{region 'Documentation'}
(*!
<summary>Number of observations from the latest subject call.</summary>
*)
{endregion}
{attribute 'monitoring' := 'call'}
PROPERTY PUBLIC HookCount : UINT //! Number of observations from the latest subject call.
GET // PUBLIC
HookCount := FHookCount;
END_GET
END_PROPERTY

{region 'Documentation'}
(*!
<summary>Combines base startability with the scenario release.</summary>
*)
{endregion}
{attribute 'monitoring' := 'call'}
PROPERTY PUBLIC IsReady : BOOL //! Combines base startability with the scenario release.
GET // PUBLIC
IsReady := SUPER^.IsReady AND Ready;
END_GET
END_PROPERTY

{region 'Documentation'}
(*!
<summary>
Records activation, supports a controlled cleanup failure and waits for the explicit completion release.
</summary>
*)
{endregion}
METHOD PROTECTED ProcessAbort
VAR_INPUT
    Enable : BOOL; //! Phase permission supplied by the owning Test Case; FALSE does not authorize progression, while observation may continue.
END_VAR
RecordHook(Hook := E_LifecycleHook.Abort,
    Enabled := Enable);
IF NOT Enable THEN
    RETURN;
END_IF;
IF AbortError THEN
    Error(Message := 'Controlled abort failure.');
END_IF;
IF AbortCompleted THEN
    CompleteAbort();
END_IF;
END_METHOD

{region 'Documentation'}
(*!
<summary>Calls both real Assertions even when disabled to consume their reset requests.</summary>
*)
{endregion}
METHOD PROTECTED ProcessAssertions
VAR_INPUT
    Enable : BOOL; //! Phase permission supplied by the owning Test Case; FALSE does not authorize progression, while observation may continue.
END_VAR
RecordHook(Hook := E_LifecycleHook.Assertions,
    Enabled := Enable);
FAssertion(Enable := Enable,
    State := State,
    IN := AssertionCondition);
FReferenceAssertion(Enable := Enable,
    State := State,
    IN := TRUE);
END_METHOD

{region 'Documentation'}
(*!
<summary>Supplies controlled target observations and explicit multi-stage completion.</summary>
*)
{endregion}
METHOD PROTECTED ProcessPreparations
VAR_INPUT
    Enable : BOOL; //! Phase permission supplied by the owning Test Case; FALSE does not authorize progression, while observation may continue.
END_VAR
RecordHook(Hook := E_LifecycleHook.Preparations,
    Enabled := Enable);
// Emulate the concrete application's combined observation without another Preparation FB.
// The Sequencer has already run; explicit completion below can still transition immediately.
UpdatePreparationStatus(Ready := TRUE,
    Running := Enable AND NOT PreparationTargetReached,
    Completed := PreparationTargetReached,
    HasError := PreparationError);
IF NOT Enable THEN
    RETURN;
END_IF;

IF AdvancePreparation THEN
    NextPreparationState();
ELSIF FinishPreparations THEN
    CompletePreparations();
END_IF;
END_METHOD

{region 'Documentation'}
(*!
<summary>Resets both real Assertions and completes only on the explicit fixture release.</summary>
*)
{endregion}
METHOD PROTECTED ProcessReset
RecordHook(Hook := E_LifecycleHook.Reset,
    Enabled := TRUE);
FAssertion.Reset();
FReferenceAssertion.Reset();
// Deliberately allow Error followed by CompleteReset in the same call.
// The base must preserve Error and choose finalization instead of a successful Idle result.
IF ResetError THEN
    Error(Message := 'Controlled reset failure.');
END_IF;
IF ResetCompleted THEN
    CompleteReset();
END_IF;
END_METHOD

{region 'Documentation'}
(*!
<summary>Advances or completes only when enabled and explicitly instructed.</summary>
*)
{endregion}
METHOD PROTECTED ProcessTests
VAR_INPUT
    Enable : BOOL; //! Phase permission supplied by the owning Test Case; FALSE does not authorize progression, while observation may continue.
END_VAR
RecordHook(Hook := E_LifecycleHook.Tests,
    Enabled := Enable);
IF NOT Enable THEN
    RETURN;
END_IF;

// Use the real base API for error and transition stimulus; never assign the subject state directly.
IF TestError THEN
    Error(Message := 'Controlled test failure.');
    RETURN;
END_IF;
IF AdvanceTest THEN
    NextTestState();
ELSIF FinishTests THEN
    CompleteTests();
END_IF;
END_METHOD

{region 'Documentation'}
(*!
<summary>Appends one hook-entry observation with bounded storage and explicit overflow reporting.</summary>
*)
{endregion}
METHOD PRIVATE RecordHook
VAR_INPUT
    Hook : E_LifecycleHook; //! Hook being entered; appended to the bounded per-call trace.
    Enabled : BOOL; //! Hook permission recorded together with the current entry state.
END_VAR
IF FHookCount >= HookCapacity THEN
    FTraceOverflow := TRUE;
    RETURN;
END_IF;

FHookCount := FHookCount + 1;
FHooks[FHookCount].Hook := Hook;
FHooks[FHookCount].State := State;
FHooks[FHookCount].Enabled := Enabled;
END_METHOD

{region 'Documentation'}
(*!
<summary>Reports a call exceeding the bounded hook trace.</summary>
*)
{endregion}
{attribute 'monitoring' := 'call'}
PROPERTY PUBLIC TraceOverflow : BOOL //! Reports a call exceeding the bounded hook trace.
GET // PUBLIC
TraceOverflow := FTraceOverflow;
END_GET
END_PROPERTY

END_FUNCTION_BLOCK

// ---- SelfTests/TestCases/TestSuite_TestCaseLifecycle/Test_LifecycleWithoutPreparation.TcPOU
{region 'Documentation'}
(*!
<summary>Checks initial passivity, parent Reset, resource readiness and explicit single-state completion.</summary>
*)
{endregion}
FUNCTION_BLOCK Test_LifecycleWithoutPreparation EXTENDS TestCaseLifecycleTestBase

SUPER^();

{region 'Documentation'}
(*!
<summary>Defines independent per-call stimuli and expected lifecycle/hook observations.</summary>
*)
{endregion}
METHOD PROTECTED ConfigureScenario
FSubjectPreparationCount := 0;
FSubjectTestCount := 1;
FStepCount := 11;

{region "01 - Initialized but awaiting Reset"}
// After successful Initialize, remain Uninitialized until the parent requests Reset.
FSteps[1].ExpectedState := E_State.Uninitialized;
FSteps[1].ExpectedResult := E_Result.NotEvaluated;
FSteps[1].ExpectedReady := FALSE;
FSteps[1].ExpectedPassedCount := 0;
FSteps[1].ExpectedFailedCount := 0;
FSteps[1].ExpectedHookCount := 5;
FSteps[1].ExpectedHooks[1].Hook := E_LifecycleHook.Abort;
FSteps[1].ExpectedHooks[1].State := E_State.Uninitialized;
FSteps[1].ExpectedHooks[1].Enabled := FALSE;
FSteps[1].ExpectedHooks[2].Hook := E_LifecycleHook.Preparations;
FSteps[1].ExpectedHooks[2].State := E_State.Uninitialized;
FSteps[1].ExpectedHooks[2].Enabled := FALSE;
FSteps[1].ExpectedHooks[3].Hook := E_LifecycleHook.Tests;
FSteps[1].ExpectedHooks[3].State := E_State.Uninitialized;
FSteps[1].ExpectedHooks[3].Enabled := FALSE;
FSteps[1].ExpectedHooks[4].Hook := E_LifecycleHook.Assertions;
FSteps[1].ExpectedHooks[4].State := E_State.Uninitialized;
FSteps[1].ExpectedHooks[4].Enabled := FALSE;
FSteps[1].ExpectedHooks[5].Hook := E_LifecycleHook.Aggregate;
FSteps[1].ExpectedHooks[5].State := E_State.Uninitialized;
FSteps[1].ExpectedHooks[5].Enabled := TRUE;
{endregion}

{region "02 - Start cannot bypass Reset"}
// Start alone must not bypass the initial Reset requirement.
FSteps[2].RequestStart := TRUE;
FSteps[2].ExpectedState := E_State.Uninitialized;
FSteps[2].ExpectedResult := E_Result.NotEvaluated;
FSteps[2].ExpectedReady := FALSE;
FSteps[2].ExpectedPassedCount := 0;
FSteps[2].ExpectedFailedCount := 0;
FSteps[2].ExpectedHookCount := 5;
FSteps[2].ExpectedHooks[1].Hook := E_LifecycleHook.Abort;
FSteps[2].ExpectedHooks[1].State := E_State.Uninitialized;
FSteps[2].ExpectedHooks[1].Enabled := FALSE;
FSteps[2].ExpectedHooks[2].Hook := E_LifecycleHook.Preparations;
FSteps[2].ExpectedHooks[2].State := E_State.Uninitialized;
FSteps[2].ExpectedHooks[2].Enabled := FALSE;
FSteps[2].ExpectedHooks[3].Hook := E_LifecycleHook.Tests;
FSteps[2].ExpectedHooks[3].State := E_State.Uninitialized;
FSteps[2].ExpectedHooks[3].Enabled := FALSE;
FSteps[2].ExpectedHooks[4].Hook := E_LifecycleHook.Assertions;
FSteps[2].ExpectedHooks[4].State := E_State.Uninitialized;
FSteps[2].ExpectedHooks[4].Enabled := FALSE;
FSteps[2].ExpectedHooks[5].Hook := E_LifecycleHook.Aggregate;
FSteps[2].ExpectedHooks[5].State := E_State.Uninitialized;
FSteps[2].ExpectedHooks[5].Enabled := TRUE;
{endregion}

{region "03 - Reset awaiting acknowledgement"}
// Accept Reset but withhold CompleteReset; the subject must remain in Reset.
FSteps[3].RequestReset := TRUE;
FSteps[3].ResetCompleted := FALSE;
FSteps[3].ExpectedState := E_State.Reset;
FSteps[3].ExpectedResult := E_Result.NotEvaluated;
FSteps[3].ExpectedReady := FALSE;
FSteps[3].ExpectedPassedCount := 0;
FSteps[3].ExpectedFailedCount := 0;
FSteps[3].ExpectedHookCount := 6;
FSteps[3].ExpectedHooks[1].Hook := E_LifecycleHook.Reset;
FSteps[3].ExpectedHooks[1].State := E_State.Reset;
FSteps[3].ExpectedHooks[1].Enabled := TRUE;
FSteps[3].ExpectedHooks[2].Hook := E_LifecycleHook.Abort;
FSteps[3].ExpectedHooks[2].State := E_State.Reset;
FSteps[3].ExpectedHooks[2].Enabled := FALSE;
FSteps[3].ExpectedHooks[3].Hook := E_LifecycleHook.Preparations;
FSteps[3].ExpectedHooks[3].State := E_State.Reset;
FSteps[3].ExpectedHooks[3].Enabled := FALSE;
FSteps[3].ExpectedHooks[4].Hook := E_LifecycleHook.Tests;
FSteps[3].ExpectedHooks[4].State := E_State.Reset;
FSteps[3].ExpectedHooks[4].Enabled := FALSE;
FSteps[3].ExpectedHooks[5].Hook := E_LifecycleHook.Assertions;
FSteps[3].ExpectedHooks[5].State := E_State.Reset;
FSteps[3].ExpectedHooks[5].Enabled := FALSE;
FSteps[3].ExpectedHooks[6].Hook := E_LifecycleHook.Aggregate;
FSteps[3].ExpectedHooks[6].State := E_State.Reset;
FSteps[3].ExpectedHooks[6].Enabled := TRUE;
{endregion}

{region "04 - Idle without readiness"}
// Release reset completion while withholding readiness: Idle does not itself imply IsReady.
FSteps[4].Ready := FALSE;
FSteps[4].ExpectedState := E_State.Idle;
FSteps[4].ExpectedResult := E_Result.NotEvaluated;
FSteps[4].ExpectedReady := FALSE;
FSteps[4].ExpectedPassedCount := 0;
FSteps[4].ExpectedFailedCount := 0;
FSteps[4].ExpectedHookCount := 6;
FSteps[4].ExpectedHooks[1].Hook := E_LifecycleHook.Reset;
FSteps[4].ExpectedHooks[1].State := E_State.Reset;
FSteps[4].ExpectedHooks[1].Enabled := TRUE;
FSteps[4].ExpectedHooks[2].Hook := E_LifecycleHook.Abort;
FSteps[4].ExpectedHooks[2].State := E_State.Idle;
FSteps[4].ExpectedHooks[2].Enabled := FALSE;
FSteps[4].ExpectedHooks[3].Hook := E_LifecycleHook.Preparations;
FSteps[4].ExpectedHooks[3].State := E_State.Idle;
FSteps[4].ExpectedHooks[3].Enabled := FALSE;
FSteps[4].ExpectedHooks[4].Hook := E_LifecycleHook.Tests;
FSteps[4].ExpectedHooks[4].State := E_State.Idle;
FSteps[4].ExpectedHooks[4].Enabled := FALSE;
FSteps[4].ExpectedHooks[5].Hook := E_LifecycleHook.Assertions;
FSteps[4].ExpectedHooks[5].State := E_State.Idle;
FSteps[4].ExpectedHooks[5].Enabled := FALSE;
FSteps[4].ExpectedHooks[6].Hook := E_LifecycleHook.Aggregate;
FSteps[4].ExpectedHooks[6].State := E_State.Idle;
FSteps[4].ExpectedHooks[6].Enabled := TRUE;
{endregion}

{region "05 - Reject Start while not ready"}
// A Start request while not ready must leave the subject in Idle.
FSteps[5].RequestStart := TRUE;
FSteps[5].Ready := FALSE;
FSteps[5].ExpectedState := E_State.Idle;
FSteps[5].ExpectedResult := E_Result.NotEvaluated;
FSteps[5].ExpectedReady := FALSE;
FSteps[5].ExpectedPassedCount := 0;
FSteps[5].ExpectedFailedCount := 0;
FSteps[5].ExpectedHookCount := 5;
FSteps[5].ExpectedHooks[1].Hook := E_LifecycleHook.Abort;
FSteps[5].ExpectedHooks[1].State := E_State.Idle;
FSteps[5].ExpectedHooks[1].Enabled := FALSE;
FSteps[5].ExpectedHooks[2].Hook := E_LifecycleHook.Preparations;
FSteps[5].ExpectedHooks[2].State := E_State.Idle;
FSteps[5].ExpectedHooks[2].Enabled := FALSE;
FSteps[5].ExpectedHooks[3].Hook := E_LifecycleHook.Tests;
FSteps[5].ExpectedHooks[3].State := E_State.Idle;
FSteps[5].ExpectedHooks[3].Enabled := FALSE;
FSteps[5].ExpectedHooks[4].Hook := E_LifecycleHook.Assertions;
FSteps[5].ExpectedHooks[4].State := E_State.Idle;
FSteps[5].ExpectedHooks[4].Enabled := FALSE;
FSteps[5].ExpectedHooks[5].Hook := E_LifecycleHook.Aggregate;
FSteps[5].ExpectedHooks[5].State := E_State.Idle;
FSteps[5].ExpectedHooks[5].Enabled := TRUE;
{endregion}

{region "06 - Ready without automatic Start"}
// Restore readiness without a fresh Start request; there must be no deferred automatic start.
FSteps[6].ExpectedState := E_State.Idle;
FSteps[6].ExpectedResult := E_Result.NotEvaluated;
FSteps[6].ExpectedReady := TRUE;
FSteps[6].ExpectedPassedCount := 0;
FSteps[6].ExpectedFailedCount := 0;
FSteps[6].ExpectedHookCount := 5;
FSteps[6].ExpectedHooks[1].Hook := E_LifecycleHook.Abort;
FSteps[6].ExpectedHooks[1].State := E_State.Idle;
FSteps[6].ExpectedHooks[1].Enabled := FALSE;
FSteps[6].ExpectedHooks[2].Hook := E_LifecycleHook.Preparations;
FSteps[6].ExpectedHooks[2].State := E_State.Idle;
FSteps[6].ExpectedHooks[2].Enabled := FALSE;
FSteps[6].ExpectedHooks[3].Hook := E_LifecycleHook.Tests;
FSteps[6].ExpectedHooks[3].State := E_State.Idle;
FSteps[6].ExpectedHooks[3].Enabled := FALSE;
FSteps[6].ExpectedHooks[4].Hook := E_LifecycleHook.Assertions;
FSteps[6].ExpectedHooks[4].State := E_State.Idle;
FSteps[6].ExpectedHooks[4].Enabled := FALSE;
FSteps[6].ExpectedHooks[5].Hook := E_LifecycleHook.Aggregate;
FSteps[6].ExpectedHooks[5].State := E_State.Idle;
FSteps[6].ExpectedHooks[5].Enabled := TRUE;
{endregion}

{region "07 - Accept fresh Start"}
// Accept Start into Starting; processing and Assertion evaluation are not active yet.
FSteps[7].RequestStart := TRUE;
FSteps[7].ExpectedState := E_State.Starting;
FSteps[7].ExpectedResult := E_Result.NotEvaluated;
FSteps[7].ExpectedReady := FALSE;
FSteps[7].ExpectedPassedCount := 0;
FSteps[7].ExpectedFailedCount := 0;
FSteps[7].ExpectedHookCount := 5;
FSteps[7].ExpectedHooks[1].Hook := E_LifecycleHook.Abort;
FSteps[7].ExpectedHooks[1].State := E_State.Starting;
FSteps[7].ExpectedHooks[1].Enabled := FALSE;
FSteps[7].ExpectedHooks[2].Hook := E_LifecycleHook.Preparations;
FSteps[7].ExpectedHooks[2].State := E_State.Starting;
FSteps[7].ExpectedHooks[2].Enabled := FALSE;
FSteps[7].ExpectedHooks[3].Hook := E_LifecycleHook.Tests;
FSteps[7].ExpectedHooks[3].State := E_State.Starting;
FSteps[7].ExpectedHooks[3].Enabled := FALSE;
FSteps[7].ExpectedHooks[4].Hook := E_LifecycleHook.Assertions;
FSteps[7].ExpectedHooks[4].State := E_State.Starting;
FSteps[7].ExpectedHooks[4].Enabled := FALSE;
FSteps[7].ExpectedHooks[5].Hook := E_LifecycleHook.Aggregate;
FSteps[7].ExpectedHooks[5].State := E_State.Starting;
FSteps[7].ExpectedHooks[5].Enabled := TRUE;
{endregion}

{region "08 - Run without Preparation"}
// Enter Running and evaluate both children; owner Result stays NotEvaluated until finalization.
FSteps[8].ExpectedState := E_State.Running;
FSteps[8].ExpectedResult := E_Result.NotEvaluated;
FSteps[8].ExpectedReady := FALSE;
FSteps[8].ExpectedPassedCount := 2;
FSteps[8].ExpectedFailedCount := 0;
FSteps[8].ExpectedHookCount := 5;
FSteps[8].ExpectedHooks[1].Hook := E_LifecycleHook.Abort;
FSteps[8].ExpectedHooks[1].State := E_State.Running;
FSteps[8].ExpectedHooks[1].Enabled := FALSE;
FSteps[8].ExpectedHooks[2].Hook := E_LifecycleHook.Preparations;
FSteps[8].ExpectedHooks[2].State := E_State.Running;
FSteps[8].ExpectedHooks[2].Enabled := FALSE;
FSteps[8].ExpectedHooks[3].Hook := E_LifecycleHook.Tests;
FSteps[8].ExpectedHooks[3].State := E_State.Running;
FSteps[8].ExpectedHooks[3].Enabled := TRUE;
FSteps[8].ExpectedHooks[4].Hook := E_LifecycleHook.Assertions;
FSteps[8].ExpectedHooks[4].State := E_State.Running;
FSteps[8].ExpectedHooks[4].Enabled := TRUE;
FSteps[8].ExpectedHooks[5].Hook := E_LifecycleHook.Aggregate;
FSteps[8].ExpectedHooks[5].State := E_State.Running;
FSteps[8].ExpectedHooks[5].Enabled := TRUE;
{endregion}

{region "09 - Keep execution open"}
// Continue Running without completion; a Passed child collection does not finish the Test Case.
FSteps[9].ExpectedState := E_State.Running;
FSteps[9].ExpectedResult := E_Result.NotEvaluated;
FSteps[9].ExpectedReady := FALSE;
FSteps[9].ExpectedPassedCount := 2;
FSteps[9].ExpectedFailedCount := 0;
FSteps[9].ExpectedHookCount := 5;
FSteps[9].ExpectedHooks[1].Hook := E_LifecycleHook.Abort;
FSteps[9].ExpectedHooks[1].State := E_State.Running;
FSteps[9].ExpectedHooks[1].Enabled := FALSE;
FSteps[9].ExpectedHooks[2].Hook := E_LifecycleHook.Preparations;
FSteps[9].ExpectedHooks[2].State := E_State.Running;
FSteps[9].ExpectedHooks[2].Enabled := FALSE;
FSteps[9].ExpectedHooks[3].Hook := E_LifecycleHook.Tests;
FSteps[9].ExpectedHooks[3].State := E_State.Running;
FSteps[9].ExpectedHooks[3].Enabled := TRUE;
FSteps[9].ExpectedHooks[4].Hook := E_LifecycleHook.Assertions;
FSteps[9].ExpectedHooks[4].State := E_State.Running;
FSteps[9].ExpectedHooks[4].Enabled := TRUE;
FSteps[9].ExpectedHooks[5].Hook := E_LifecycleHook.Aggregate;
FSteps[9].ExpectedHooks[5].State := E_State.Running;
FSteps[9].ExpectedHooks[5].Enabled := TRUE;
{endregion}

{region "10 - Complete inside test processing"}
// CompleteTests changes phase inside ProcessTests; subsequent Assertions must already be
// disabled.
FSteps[10].FinishTests := TRUE;
FSteps[10].ExpectedState := E_State.Completing;
FSteps[10].ExpectedResult := E_Result.Passed;
FSteps[10].ExpectedReady := FALSE;
FSteps[10].ExpectedPassedCount := 2;
FSteps[10].ExpectedFailedCount := 0;
FSteps[10].ExpectedHookCount := 5;
FSteps[10].ExpectedHooks[1].Hook := E_LifecycleHook.Abort;
FSteps[10].ExpectedHooks[1].State := E_State.Running;
FSteps[10].ExpectedHooks[1].Enabled := FALSE;
FSteps[10].ExpectedHooks[2].Hook := E_LifecycleHook.Preparations;
FSteps[10].ExpectedHooks[2].State := E_State.Running;
FSteps[10].ExpectedHooks[2].Enabled := FALSE;
FSteps[10].ExpectedHooks[3].Hook := E_LifecycleHook.Tests;
FSteps[10].ExpectedHooks[3].State := E_State.Running;
FSteps[10].ExpectedHooks[3].Enabled := TRUE;
FSteps[10].ExpectedHooks[4].Hook := E_LifecycleHook.Assertions;
FSteps[10].ExpectedHooks[4].State := E_State.Completing;
FSteps[10].ExpectedHooks[4].Enabled := FALSE;
FSteps[10].ExpectedHooks[5].Hook := E_LifecycleHook.Aggregate;
FSteps[10].ExpectedHooks[5].State := E_State.Completing;
FSteps[10].ExpectedHooks[5].Enabled := TRUE;
{endregion}

{region "11 - Observe terminal completion"}
// The following call reaches Completed; only aggregation remains in the recorded processing
// hooks.
FSteps[11].ExpectedState := E_State.Completed;
FSteps[11].ExpectedResult := E_Result.Passed;
FSteps[11].ExpectedReady := FALSE;
FSteps[11].ExpectedPassedCount := 2;
FSteps[11].ExpectedFailedCount := 0;
FSteps[11].ExpectedHookCount := 1;
FSteps[11].ExpectedHooks[1].Hook := E_LifecycleHook.Aggregate;
FSteps[11].ExpectedHooks[1].State := E_State.Completed;
FSteps[11].ExpectedHooks[1].Enabled := TRUE;
{endregion}
END_METHOD

END_FUNCTION_BLOCK

// ---- SelfTests/TestCases/TestSuite_TestCaseLifecycle/Helper/TestCaseLifecycleTestBase.TcPOU
{region 'Documentation'}
(*!
<summary>
Drives and checks an isolated TestCaseBase-derived subject using explicit scenario checkpoints.
</summary>

<description>

Roles and isolation

The outer Test Case is the selftest; FSubject is the object under test.

FSubject executes the real inherited lifecycle, not a copied Sequencer.

Subject and child-Assertion events remain in FCapture.

Outer checking Assertions report through the regular framework publisher.

An expected subject Failed or Error result can therefore pass the outer selftest.
BindSubjectParent supplies the containing Suite identity; only this test calls FSubject.

Scenario checkpoints

ConfigureScenario supplies FSteps with stimuli and independent expectations.
A step is a checkpoint, not a subject lifecycle state.
ProcessTests applies the stimuli and calls the subject once per active cycle.
ProcessAssertions checks the resulting status and trace before the next step starts.
Waiting checkpoints may span several PLC cycles without blocking the task.

Hook observations

The subject records each Process* and AggregateResults method entry:
method, current state and received Enable.
The trace covers one subject call and is separate from event logging.
Comparing these entries tests the agreed call order, including state changes
between two hooks in the same call.

Terminal and repeat-run evidence

Optional event checkpoints count Result, Aggregation and Completed transitions in the
isolated capture. No entries are deleted; a subject Reset retains earlier event evidence.
Quiet-call checks reject any new event; runtime checks distinguish clearing from holding.
</description>
*)
{endregion}
FUNCTION_BLOCK ABSTRACT TestCaseLifecycleTestBase EXTENDS TestCaseBase
VAR
    FSteps : ARRAY[1..StepCapacity] OF ST_LifecycleStep;
    FStepCount : INT;
    FSubjectPreparationCount : INT;
    FSubjectTestCount : INT;
    FSubjectParent : I_TestSuite;
    FSubject : TestCaseLifecycleProbe;
    FCapture : EventBuffer;
    FEvents : ARRAY[1..CaptureLength] OF ST_Event;
    FCaptureFifo : ST_FifoStatus;
    FCaptureStatus : ST_EventBufferStatus;
    FFixtureValid : BOOL;
    FStepIndex : INT := 1;
    FCheckPerformed : BOOL;
    FObserved : ST_TestCaseStatus;
    FHookOrderMatches : BOOL;
    FHookStatesMatch : BOOL;
    FHookEnableMatches : BOOL;
    FCheckState : AssertEqual_Int;
    FCheckResult : AssertEqual_Int;
    FCheckReady : AssertEqual_Bool;
    FCheckStatusReady : AssertEqual_Bool;
    FCheckTotalCount : AssertEqual_UInt;
    FCheckPassedCount : AssertEqual_UInt;
    FCheckFailedCount : AssertEqual_UInt;
    FCheckHookCount : AssertEqual_UInt;
    FCheckHookOrder : AssertTrue;
    FCheckHookStates : AssertTrue;
    FCheckHookEnable : AssertTrue;
    FCheckTraceBound : AssertFalse;
    FCheckNoLostEvents : AssertEqual_UDInt;
    FSubjectConfig : ST_TestCaseConfig;
    FObservationReady : BOOL;
    FCheckHasError : AssertEqual_Bool;
    FCheckStatusError : AssertEqual_Bool;
    FCheckTimeout : AssertEqual_Bool;
    FCheckPreparationTimeout : AssertEqual_Bool;
    FCheckResetTimeout : AssertEqual_Bool;
    FCheckAbortTimeout : AssertEqual_Bool;
    FPreviousRuntime : TIME;
    FSequenceBeforeCall : UDINT;
    FCheckFinalization : AssertTrue;
    FCheckQuietCall : AssertTrue;
    FCheckRuntime : AssertTrue;
    FCheckStatusProjection : AssertTrue;
END_VAR
VAR CONSTANT
    StepCapacity : INT := 24;
    CaptureLength : UINT := 256;
END_VAR

SUPER^();

{region 'Documentation'}
(*!
<summary>Contributes every outer Assertion once without advancing the fixture.</summary>
*)
{endregion}
METHOD PROTECTED AggregateResults
VAR_INPUT
    Aggregator : I_ResultAggregator; //! Borrowed result sink owned by the outer Test Case; add this test's checking Assertions without resetting or retaining the sink.
END_VAR
Aggregator.AddProvider(Provider := FCheckState);
Aggregator.AddProvider(Provider := FCheckResult);
Aggregator.AddProvider(Provider := FCheckReady);
Aggregator.AddProvider(Provider := FCheckStatusReady);
Aggregator.AddProvider(Provider := FCheckTotalCount);
Aggregator.AddProvider(Provider := FCheckPassedCount);
Aggregator.AddProvider(Provider := FCheckFailedCount);
Aggregator.AddProvider(Provider := FCheckHookCount);
Aggregator.AddProvider(Provider := FCheckHookOrder);
Aggregator.AddProvider(Provider := FCheckHookStates);
Aggregator.AddProvider(Provider := FCheckHookEnable);
Aggregator.AddProvider(Provider := FCheckTraceBound);
Aggregator.AddProvider(Provider := FCheckNoLostEvents);
Aggregator.AddProvider(Provider := FCheckHasError);
Aggregator.AddProvider(Provider := FCheckStatusError);
Aggregator.AddProvider(Provider := FCheckTimeout);
Aggregator.AddProvider(Provider := FCheckPreparationTimeout);
Aggregator.AddProvider(Provider := FCheckResetTimeout);
Aggregator.AddProvider(Provider := FCheckAbortTimeout);
Aggregator.AddProvider(Provider := FCheckFinalization);
Aggregator.AddProvider(Provider := FCheckQuietCall);
Aggregator.AddProvider(Provider := FCheckRuntime);
Aggregator.AddProvider(Provider := FCheckStatusProjection);
END_METHOD

{region 'Documentation'}
(*!
<summary>Checks retained finalization evidence against this checkpoint, without deriving expected counts from the subject.</summary>
<description>
The local capture is never consumed or overwritten within a scenario. Entries therefore
remain in publication order from index 1. The guard rejects loss or an unexpected layout.
Only this subject's owner events count; Assertion findings remain separate evidence.
Each Result must be followed by one Aggregation in Completing and then a Completed transition.
</description>
*)
{endregion}
METHOD PRIVATE AreFinalizationEventsValid : BOOL //! TRUE when finalization checking is disabled or the retained ordered owner events match this checkpoint.
VAR
    Index : UINT;
    Event : REFERENCE TO ST_Event;
    ResultCount : UINT;
    AggregationCount : UINT;
    CompletionCount : UINT;
    LastResult : E_Result;
    PreviousSequence : UDINT;
END_VAR
AreFinalizationEventsValid := TRUE;
IF NOT FSteps[FStepIndex].CheckFinalization THEN
    RETURN;
END_IF;
AreFinalizationEventsValid := FALSE;
IF FCaptureFifo.ConfigError OR FCaptureFifo.IndexError
    OR (FCaptureStatus.LostEventCount <> 0)
    OR (FCaptureFifo.ElementCount >= CaptureLength)
    OR (FCaptureFifo.IndexOut <> 1)
    OR (FCaptureStatus.SequenceId <> UINT_TO_UDINT(FCaptureFifo.ElementCount)) THEN
    RETURN;
END_IF;

FOR Index := 1 TO FCaptureFifo.ElementCount DO
    Event REF= FEvents[Index];
    IF Event.SequenceId <= PreviousSequence THEN
        RETURN;
    END_IF;
    PreviousSequence := Event.SequenceId;
    IF (Event.OwnerScope <> E_OwnerScope.TestCase) OR (Event.Name <> FSubject.Name) THEN
        CONTINUE;
    END_IF;

    CASE Event.EventType OF
        E_EventType.Result:
            IF (Event.State <> E_State.Completing)
                OR (ResultCount <> CompletionCount) OR (AggregationCount <> CompletionCount) THEN
                RETURN;
            END_IF;
            ResultCount := ResultCount + 1;
            LastResult := Event.Result;

        E_EventType.Aggregation:
            IF (Event.State <> E_State.Completing) OR (Event.Result <> LastResult)
                OR (ResultCount <> AggregationCount + 1) OR (AggregationCount <> CompletionCount) THEN
                RETURN;
            END_IF;
            AggregationCount := AggregationCount + 1;

        E_EventType.StateTransition:
            IF Event.State = E_State.Completed THEN
                IF (ResultCount <> CompletionCount + 1) OR (AggregationCount <> ResultCount) THEN
                    RETURN;
                END_IF;
                CompletionCount := CompletionCount + 1;
            END_IF;
    ELSE
        // Triggers and technical diagnostics do not finalize the owner.
        CONTINUE;
    END_CASE;
END_FOR;

IF (ResultCount <> FSteps[FStepIndex].ExpectedFinalizationCount)
    OR (AggregationCount <> FSteps[FStepIndex].ExpectedFinalizationCount)
    OR (CompletionCount <> FSteps[FStepIndex].ExpectedCompletionCount) THEN
    RETURN;
END_IF;
IF (ResultCount > 0) AND (LastResult <> FSteps[FStepIndex].ExpectedFinalResult) THEN
    RETURN;
END_IF;

AreFinalizationEventsValid := TRUE;
END_METHOD

{region 'Documentation'}
(*!
<summary>Supplies the real containing Suite identity before this outer Test Case is initialized.</summary>
*)
{endregion}
METHOD PUBLIC BindSubjectParent
VAR_INPUT
    Parent : I_TestSuite; //! Borrowed identity parent retained for isolated subject initialization; keep the Suite alive through subject use.
END_VAR
FSubjectParent := Parent;
END_METHOD

{region 'Documentation'}
(*!
<summary>Requires a complete cycle table, a valid fixture and all evaluating Assertions.</summary>
*)
{endregion}
METHOD PROTECTED CheckInitialization : BOOL //! TRUE when the inherited initialization check and this concrete fixture check both accept the setup.

VAR
    Index : INT;
END_VAR
CheckInitialization := FALSE;
IF NOT SUPER^.CheckInitialization() THEN
    RETURN;
END_IF;
IF (FStepCount < 1) OR (FStepCount > StepCapacity) OR NOT FFixtureValid THEN
    RETURN;
END_IF;
IF NOT FCheckState.IsInitialized
    OR NOT FCheckResult.IsInitialized
    OR NOT FCheckReady.IsInitialized
    OR NOT FCheckStatusReady.IsInitialized
    OR NOT FCheckTotalCount.IsInitialized
    OR NOT FCheckPassedCount.IsInitialized
    OR NOT FCheckFailedCount.IsInitialized
    OR NOT FCheckHookCount.IsInitialized
    OR NOT FCheckHookOrder.IsInitialized
    OR NOT FCheckHookStates.IsInitialized
    OR NOT FCheckHookEnable.IsInitialized
    OR NOT FCheckTraceBound.IsInitialized
    OR NOT FCheckNoLostEvents.IsInitialized
    OR NOT FCheckHasError.IsInitialized
    OR NOT FCheckStatusError.IsInitialized
    OR NOT FCheckTimeout.IsInitialized
    OR NOT FCheckPreparationTimeout.IsInitialized
    OR NOT FCheckResetTimeout.IsInitialized
    OR NOT FCheckAbortTimeout.IsInitialized
    OR NOT FCheckFinalization.IsInitialized
    OR NOT FCheckQuietCall.IsInitialized
    OR NOT FCheckRuntime.IsInitialized
    OR NOT FCheckStatusProjection.IsInitialized THEN
    RETURN;
END_IF;

FOR Index := 1 TO FStepCount DO
    IF (FSteps[Index].ExpectedHookCount < 1)
        OR (FSteps[Index].ExpectedHookCount > 6) THEN
        RETURN;
    END_IF;
END_FOR;

CheckInitialization := TRUE;
END_METHOD

{region 'Documentation'}
(*!
<summary>Compares the bounded trace with independently authored hook order, state and enable expectations.</summary>
*)
{endregion}
METHOD PRIVATE CompareHookTrace
VAR
    Index : UINT;
    Observed : ST_LifecycleHook;
END_VAR
// Compare against the scenario's explicit trace, never against an expectation derived from FSubject.
// Count is checked separately so extra calls cannot pass just because the expected prefix matches.
FHookOrderMatches := TRUE;
FHookStatesMatch := TRUE;
FHookEnableMatches := TRUE;
FOR Index := 1 TO FSteps[FStepIndex].ExpectedHookCount DO
    Observed := FSubject.GetHook(Index := Index);
    FHookOrderMatches := FHookOrderMatches AND (Observed.Hook = FSteps[FStepIndex].ExpectedHooks[Index].Hook);
    FHookStatesMatch := FHookStatesMatch AND (Observed.State = FSteps[FStepIndex].ExpectedHooks[Index].State);
    FHookEnableMatches := FHookEnableMatches AND (Observed.Enabled = FSteps[FStepIndex].ExpectedHooks[Index].Enabled);
END_FOR;
END_METHOD

{region 'Documentation'}
(*!
<summary>Defines the scenario, initializes isolated capture and names the evaluating Assertions.</summary>
*)
{endregion}
METHOD PROTECTED Configure
VAR
    Index : INT;
    EmptyStep : ST_LifecycleStep;
    DefaultConfig : ST_TestCaseConfig;
END_VAR
// Each row starts independently from the DUT defaults, not from the preceding row.
FOR Index := 1 TO StepCapacity DO
    FSteps[Index] := EmptyStep;
END_FOR;
FStepCount := 0;
FSubjectPreparationCount := 0;
FSubjectTestCount := 1;
FSubjectConfig := DefaultConfig;
ConfigureScenario();
// Outer Test states identify checkpoints; subject state counts belong to the separate fixture.
FPreparationStateCount := 0;
FTestStateCount := FStepCount;
FStepIndex := 1;
FCheckPerformed := FALSE;
FObservationReady := FALSE;
FFixtureValid := InitializeSubject();

// These Assertions judge the subject and report through the regular selftest publisher.
FCheckState.Initialize(Parent := THIS^,
    AssertionName := 'State');
FCheckResult.Initialize(Parent := THIS^,
    AssertionName := 'Result');
FCheckReady.Initialize(Parent := THIS^,
    AssertionName := 'Ready');
FCheckStatusReady.Initialize(Parent := THIS^,
    AssertionName := 'StatusReady');
FCheckTotalCount.Initialize(Parent := THIS^,
    AssertionName := 'TotalCount');
FCheckPassedCount.Initialize(Parent := THIS^,
    AssertionName := 'PassedCount');
FCheckFailedCount.Initialize(Parent := THIS^,
    AssertionName := 'FailedCount');
FCheckHookCount.Initialize(Parent := THIS^,
    AssertionName := 'HookCount');
FCheckHookOrder.Initialize(Parent := THIS^,
    AssertionName := 'HookOrder');
FCheckHookStates.Initialize(Parent := THIS^,
    AssertionName := 'HookStates');
FCheckHookEnable.Initialize(Parent := THIS^,
    AssertionName := 'HookEnable');
FCheckTraceBound.Initialize(Parent := THIS^,
    AssertionName := 'TraceBound');
FCheckNoLostEvents.Initialize(Parent := THIS^,
    AssertionName := 'NoLostEvents');
FCheckHasError.Initialize(Parent := THIS^,
    AssertionName := 'HasError');
FCheckStatusError.Initialize(Parent := THIS^,
    AssertionName := 'StatusError');
FCheckTimeout.Initialize(Parent := THIS^,
    AssertionName := 'Timeout');
FCheckPreparationTimeout.Initialize(Parent := THIS^,
    AssertionName := 'PreparationTimeout');
FCheckResetTimeout.Initialize(Parent := THIS^,
    AssertionName := 'ResetTimeout');
FCheckAbortTimeout.Initialize(Parent := THIS^,
    AssertionName := 'AbortTimeout');
FCheckFinalization.Initialize(Parent := THIS^,
    AssertionName := 'Finalization');
FCheckQuietCall.Initialize(Parent := THIS^,
    AssertionName := 'QuietCall');
FCheckRuntime.Initialize(Parent := THIS^,
    AssertionName := 'Runtime');
FCheckStatusProjection.Initialize(Parent := THIS^,
    AssertionName := 'StatusProjection');
END_METHOD

{region 'Documentation'}
(*!
<summary>Defines phase counts and a bounded, explicit stimulus/expectation table.</summary>
*)
{endregion}
METHOD PROTECTED ABSTRACT ConfigureScenario
END_METHOD

{region 'Documentation'}
(*!
<summary>Rebuilds only the isolated fixture with a fresh buffer and the agreed pre-use binding.</summary>
*)
{endregion}
METHOD PRIVATE InitializeSubject : BOOL //! TRUE when isolated capture and controlled Test Case initialization both succeed.
InitializeSubject := FALSE;
IF NOT FCapture.Initialize(Buffer := FEvents,
    FifoControl := FCaptureFifo,
    Status := FCaptureStatus) THEN
    RETURN;
END_IF;

// Bind before Initialize: even initialization diagnostics must stay in the local capture.
// The Suite supplies identity only; the subject is driven exclusively by this outer test.
FSubject.Bind(Publisher := FCapture,
    PreparationCount := FSubjectPreparationCount,
    TestCount := FSubjectTestCount);
InitializeSubject := FSubject.Initialize(Parent := FSubjectParent,
    TestName := 'Subject',
    Config := FSubjectConfig);
END_METHOD

{region 'Documentation'}
(*!
<summary>Stops invoking the local subject; it owns no external resource.</summary>
*)
{endregion}
METHOD PROTECTED ProcessAbort
VAR_INPUT
    Enable : BOOL; //! Phase permission supplied by the owning Test Case; FALSE does not authorize progression, while observation may continue.
END_VAR
IF Enable THEN
    CompleteAbort();
END_IF;
END_METHOD

{region 'Documentation'}
(*!
<summary>Evaluates the captured lifecycle and trace; disabled calls still consume pending Assertion resets.</summary>
*)
{endregion}
METHOD PROTECTED ProcessAssertions
VAR_INPUT
    Enable : BOOL; //! Phase permission supplied by the owning Test Case; FALSE does not authorize progression, while observation may continue.
END_VAR
VAR
    EvaluateChecks : BOOL;
END_VAR
// A waiting row has no final observation yet. Still call the Assertions disabled
// so pending Assertion resets are processed through their normal cyclic path.
EvaluateChecks := Enable AND FObservationReady;

FCheckState(Enable := EvaluateChecks,
    State := State,
    IN := TO_INT(FSubject.State),
    Expected := TO_INT(FSteps[FStepIndex].ExpectedState));
FCheckResult(Enable := EvaluateChecks,
    State := State,
    IN := TO_INT(FSubject.Result),
    Expected := TO_INT(FSteps[FStepIndex].ExpectedResult));
FCheckReady(Enable := EvaluateChecks,
    State := State,
    IN := FSubject.IsReady,
    Expected := FSteps[FStepIndex].ExpectedReady);
FCheckStatusReady(Enable := EvaluateChecks,
    State := State,
    IN := FObserved.Execution.Ready,
    Expected := FSteps[FStepIndex].ExpectedReady);
FCheckTotalCount(Enable := EvaluateChecks,
    State := State,
    IN := FObserved.AssertionCountTotal,
    Expected := 2);
FCheckPassedCount(Enable := EvaluateChecks,
    State := State,
    IN := FObserved.AssertionCountPassed,
    Expected := FSteps[FStepIndex].ExpectedPassedCount);
FCheckFailedCount(Enable := EvaluateChecks,
    State := State,
    IN := FObserved.AssertionCountFailed,
    Expected := FSteps[FStepIndex].ExpectedFailedCount);
FCheckHookCount(Enable := EvaluateChecks,
    State := State,
    IN := FSubject.HookCount,
    Expected := FSteps[FStepIndex].ExpectedHookCount);
FCheckHookOrder(Enable := EvaluateChecks,
    State := State,
    IN := FHookOrderMatches);
FCheckHookStates(Enable := EvaluateChecks,
    State := State,
    IN := FHookStatesMatch);
FCheckHookEnable(Enable := EvaluateChecks,
    State := State,
    IN := FHookEnableMatches);
FCheckTraceBound(Enable := EvaluateChecks,
    State := State,
    IN := FSubject.TraceOverflow);
FCheckNoLostEvents(Enable := EvaluateChecks,
    State := State,
    IN := FCaptureStatus.LostEventCount,
    Expected := 0);
FCheckHasError(Enable := EvaluateChecks,
    State := State,
    IN := FSubject.HasError,
    Expected := FSteps[FStepIndex].ExpectedResult = E_Result.Error);
FCheckStatusError(Enable := EvaluateChecks,
    State := State,
    IN := FObserved.Execution.Error,
    Expected := FSteps[FStepIndex].ExpectedResult = E_Result.Error);
FCheckTimeout(Enable := EvaluateChecks,
    State := State,
    IN := FSubject.HasTimeout,
    Expected := FSteps[FStepIndex].ExpectedTimeout);
FCheckPreparationTimeout(Enable := EvaluateChecks,
    State := State,
    IN := FSubject.HasPreparationTimeout,
    Expected := FSteps[FStepIndex].ExpectedPreparationTimeout);
FCheckResetTimeout(Enable := EvaluateChecks,
    State := State,
    IN := FSubject.HasResetTimeout,
    Expected := FSteps[FStepIndex].ExpectedResetTimeout);
FCheckAbortTimeout(Enable := EvaluateChecks,
    State := State,
    IN := FSubject.HasAbortTimeout,
    Expected := FSteps[FStepIndex].ExpectedAbortTimeout);

FCheckFinalization(Enable := EvaluateChecks,
    State := State,
    IN := AreFinalizationEventsValid());
FCheckQuietCall(Enable := EvaluateChecks,
    State := State,
    IN := NOT FSteps[FStepIndex].ExpectQuietCall
        OR (FCaptureStatus.SequenceId = FSequenceBeforeCall));
FCheckRuntime(Enable := EvaluateChecks,
    State := State,
    IN := (NOT FSteps[FStepIndex].ExpectRuntimeCleared OR (FObserved.Runtime = T#0ms))
        AND (NOT FSteps[FStepIndex].ExpectRuntimeHeld OR (FObserved.Runtime = FPreviousRuntime)));
FCheckStatusProjection(Enable := EvaluateChecks,
    State := State,
    IN := (FObserved.Execution.State = FSteps[FStepIndex].ExpectedState)
        AND (FObserved.Execution.Result = FSteps[FStepIndex].ExpectedResult)
        AND (FObserved.Execution.Completed = (FSteps[FStepIndex].ExpectedState = E_State.Completed))
        AND (FObserved.Execution.Uninitialized = (FSteps[FStepIndex].ExpectedState = E_State.Uninitialized))
        AND (FObserved.Execution.Aborted = ((FSteps[FStepIndex].ExpectedState = E_State.Completed)
            AND (FSteps[FStepIndex].ExpectedResult = E_Result.Abort)))
        AND NOT FObserved.Execution.ConfigError);

// Do not advance merely because checks were called: their evaluation gate must be active.
// Results remain latched across checkpoints, so a later matching row cannot hide a failure.
IF EvaluateChecks
    AND FCheckState.EvaluationActive
    AND FCheckResult.EvaluationActive
    AND FCheckReady.EvaluationActive
    AND FCheckStatusReady.EvaluationActive
    AND FCheckTotalCount.EvaluationActive
    AND FCheckPassedCount.EvaluationActive
    AND FCheckFailedCount.EvaluationActive
    AND FCheckHookCount.EvaluationActive
    AND FCheckHookOrder.EvaluationActive
    AND FCheckHookStates.EvaluationActive
    AND FCheckHookEnable.EvaluationActive
    AND FCheckTraceBound.EvaluationActive
    AND FCheckNoLostEvents.EvaluationActive
    AND FCheckHasError.EvaluationActive
    AND FCheckStatusError.EvaluationActive
    AND FCheckTimeout.EvaluationActive
    AND FCheckPreparationTimeout.EvaluationActive
    AND FCheckResetTimeout.EvaluationActive
    AND FCheckAbortTimeout.EvaluationActive
    AND FCheckFinalization.EvaluationActive
    AND FCheckQuietCall.EvaluationActive
    AND FCheckRuntime.EvaluationActive
    AND FCheckStatusProjection.EvaluationActive THEN
    FCheckPerformed := TRUE;
END_IF;
END_METHOD

{region 'Documentation'}
(*!
<summary>No outer Preparation phase is needed; subject Preparation is test stimulus.</summary>
*)
{endregion}
METHOD PROTECTED ProcessPreparations
VAR_INPUT
    // SA0033: Required hook without an outer Preparation phase.
    {attribute 'analysis' := '-33'}
    Enable : BOOL; //! Phase permission supplied by the owning Test Case; FALSE does not authorize progression, while observation may continue.
END_VAR
END_METHOD

{region 'Documentation'}
(*!
<summary>Reinitializes the isolated subject/capture and clears outer Assertion results for repeatable runs.</summary>
*)
{endregion}
METHOD PROTECTED ProcessReset
FStepIndex := 1;
FCheckPerformed := FALSE;
FObservationReady := FALSE;
FCheckState.Reset();
FCheckResult.Reset();
FCheckReady.Reset();
FCheckStatusReady.Reset();
FCheckTotalCount.Reset();
FCheckPassedCount.Reset();
FCheckFailedCount.Reset();
FCheckHookCount.Reset();
FCheckHookOrder.Reset();
FCheckHookStates.Reset();
FCheckHookEnable.Reset();
FCheckTraceBound.Reset();
FCheckNoLostEvents.Reset();
FCheckHasError.Reset();
FCheckStatusError.Reset();
FCheckTimeout.Reset();
FCheckPreparationTimeout.Reset();
FCheckResetTimeout.Reset();
FCheckAbortTimeout.Reset();
FCheckFinalization.Reset();
FCheckQuietCall.Reset();
FCheckRuntime.Reset();
FCheckStatusProjection.Reset();
// Reset of the OUTER test rebuilds its fixture for repeatability.
// Reset of the SUBJECT is a separate scenario stimulus in FSteps, not this setup operation.
FFixtureValid := InitializeSubject();
IF NOT FFixtureValid THEN
    Error(Message := 'Lifecycle subject setup failed.');
END_IF;
CompleteReset();
END_METHOD

{region 'Documentation'}
(*!
<summary>Executes exactly one subject call per active outer cycle and checks every step before advancing.</summary>
*)
{endregion}
METHOD PROTECTED ProcessTests
VAR_INPUT
    Enable : BOOL; //! Phase permission supplied by the owning Test Case; FALSE does not authorize progression, while observation may continue.
END_VAR
IF NOT Enable THEN
    RETURN;
END_IF;

// Advance only after ProcessAssertions evaluated the previous checkpoint.
// A failed check is retained by the outer Assertion; evaluation does not imply success.
FObservationReady := FALSE;
IF FCheckPerformed THEN
    FCheckPerformed := FALSE;
    IF FStepIndex = FStepCount THEN
        CompleteTests();
        RETURN;
    END_IF;
    FStepIndex := FStepIndex + 1;
    NextTestState();
    IF NOT IsTestingActive THEN
        RETURN;
    END_IF;
END_IF;

// Act as the subject's owner: reserve first, then submit the row's one-shot requests.
// Request priority itself is exercised by the subject, not preselected by this driver.
IF FSteps[FStepIndex].RequestReset THEN
    IF FSubject.ReserveResetEvents() <> E_EventReservationResult.Accepted THEN
        Error(Message := 'Lifecycle fixture could not reserve Reset events.');
        RETURN;
    END_IF;
    FSubject.RequestReset();
END_IF;
IF FSteps[FStepIndex].RequestStart THEN
    IF FSubject.ReserveExecutionEvents() <> E_EventReservationResult.Accepted THEN
        Error(Message := 'Lifecycle fixture could not reserve execution events.');
        RETURN;
    END_IF;
    FSubject.RequestStart();
END_IF;

IF FSteps[FStepIndex].RequestAbort THEN
    FSubject.RequestAbort();
END_IF;

FPreviousRuntime := FObserved.Runtime;
FSequenceBeforeCall := FCaptureStatus.SequenceId;

// One synchronous subject call produces the status and hook trace for this checkpoint.
FSubject(Ready := FSteps[FStepIndex].Ready,
    ResetCompleted := FSteps[FStepIndex].ResetCompleted,
    PreparationTargetReached := FSteps[FStepIndex].PreparationTargetReached,
    AdvancePreparation := FSteps[FStepIndex].AdvancePreparation,
    FinishPreparations := FSteps[FStepIndex].FinishPreparations,
    AdvanceTest := FSteps[FStepIndex].AdvanceTest,
    FinishTests := FSteps[FStepIndex].FinishTests,
    AssertionCondition := FSteps[FStepIndex].AssertionCondition,
    AbortCompleted := FSteps[FStepIndex].AbortCompleted,
    ResetError := FSteps[FStepIndex].ResetError,
    TestError := FSteps[FStepIndex].TestError,
    AbortError := FSteps[FStepIndex].AbortError,
    PreparationError := FSteps[FStepIndex].PreparationError);
FObserved := FSubject.Status;
// Timeout scenarios keep calling once per cycle, without reissuing the preceding request.
// Any state other than WaitingState is checked below, including an unexpected transition.
IF FSteps[FStepIndex].WaitForTransition
    AND (FSubject.State = FSteps[FStepIndex].WaitingState) THEN
    RETURN;
END_IF;

// The following ProcessAssertions call may now evaluate this observation.
FObservationReady := TRUE;
CompareHookTrace();
// Release the local reservation at a stable boundary, but retain captured events.
IF FSubject.IsReady OR FSubject.IsComplete THEN
    IF NOT FSubject.FreeReservedEvents() THEN
        Error(Message := 'Lifecycle fixture could not release its reservation.');
    END_IF;
END_IF;
END_METHOD

END_FUNCTION_BLOCK

// ---- Framework/Assertions/POU/BasicTypes/Bool/AssertFalse.TcPOU
{region 'Documentation'}
(*!
<summary>Checks that the BOOL value is FALSE.</summary>
*)
{endregion}
FUNCTION_BLOCK AssertFalse EXTENDS AssertionBase
VAR_INPUT
    IN : BOOL; //! Actual value checked or observed by this Assertion.
END_VAR

SUPER^();

{region 'Documentation'}
(*!
<summary>Evaluate whether the BOOL value is FALSE.</summary>
*)
{endregion}
METHOD PROTECTED Assert
VAR
    Message : STRING(GVL_Constants.MessageLength);
    ActualText : STRING(GVL_Constants.AssertionValueLength);
END_VAR
IF NOT EvaluationActive THEN
    RETURN;
END_IF;

IF Result = E_Result.Error THEN
    RETURN;
END_IF;

IF Result = E_Result.Failed THEN
    RETURN;
END_IF;

IF IN THEN
    ActualText := BOOL_TO_STRING(IN);
    Message := CONCAT('Assertion failed: values are not equal. Expected = FALSE, Actual = ',
        ActualText);
    Message := CONCAT(Message, '.');
    Fail(Message := Message);
    RETURN;
END_IF;

Pass();
END_METHOD

END_FUNCTION_BLOCK

// ---- SelfTests/TestCases/TestSuite_TestCaseLifecycle/Test_LifecycleSinglePreparation.TcPOU
{region 'Documentation'}
(*!
<summary>Checks a pending target, observation-driven handover and one explicit Test state.</summary>
*)
{endregion}
FUNCTION_BLOCK Test_LifecycleSinglePreparation EXTENDS TestCaseLifecycleTestBase

SUPER^();

{region 'Documentation'}
(*!
<summary>Defines independent per-call stimuli and expected lifecycle/hook observations.</summary>
*)
{endregion}
METHOD PROTECTED ConfigureScenario
FSubjectPreparationCount := 1;
FSubjectTestCount := 1;
FStepCount := 7;

{region "01 - Reset to Idle"}
// Establish Idle through the parent Reset request; both child results must be cleared.
FSteps[1].RequestReset := TRUE;
FSteps[1].ExpectedState := E_State.Idle;
FSteps[1].ExpectedResult := E_Result.NotEvaluated;
FSteps[1].ExpectedReady := TRUE;
FSteps[1].ExpectedPassedCount := 0;
FSteps[1].ExpectedFailedCount := 0;
FSteps[1].ExpectedHookCount := 6;
FSteps[1].ExpectedHooks[1].Hook := E_LifecycleHook.Reset;
FSteps[1].ExpectedHooks[1].State := E_State.Reset;
FSteps[1].ExpectedHooks[1].Enabled := TRUE;
FSteps[1].ExpectedHooks[2].Hook := E_LifecycleHook.Abort;
FSteps[1].ExpectedHooks[2].State := E_State.Idle;
FSteps[1].ExpectedHooks[2].Enabled := FALSE;
FSteps[1].ExpectedHooks[3].Hook := E_LifecycleHook.Preparations;
FSteps[1].ExpectedHooks[3].State := E_State.Idle;
FSteps[1].ExpectedHooks[3].Enabled := FALSE;
FSteps[1].ExpectedHooks[4].Hook := E_LifecycleHook.Tests;
FSteps[1].ExpectedHooks[4].State := E_State.Idle;
FSteps[1].ExpectedHooks[4].Enabled := FALSE;
FSteps[1].ExpectedHooks[5].Hook := E_LifecycleHook.Assertions;
FSteps[1].ExpectedHooks[5].State := E_State.Idle;
FSteps[1].ExpectedHooks[5].Enabled := FALSE;
FSteps[1].ExpectedHooks[6].Hook := E_LifecycleHook.Aggregate;
FSteps[1].ExpectedHooks[6].State := E_State.Idle;
FSteps[1].ExpectedHooks[6].Enabled := TRUE;
{endregion}

{region "02 - Accept Start"}
// Accept Start into Starting; processing and Assertion evaluation are not active yet.
FSteps[2].RequestStart := TRUE;
FSteps[2].ExpectedState := E_State.Starting;
FSteps[2].ExpectedResult := E_Result.NotEvaluated;
FSteps[2].ExpectedReady := FALSE;
FSteps[2].ExpectedPassedCount := 0;
FSteps[2].ExpectedFailedCount := 0;
FSteps[2].ExpectedHookCount := 5;
FSteps[2].ExpectedHooks[1].Hook := E_LifecycleHook.Abort;
FSteps[2].ExpectedHooks[1].State := E_State.Starting;
FSteps[2].ExpectedHooks[1].Enabled := FALSE;
FSteps[2].ExpectedHooks[2].Hook := E_LifecycleHook.Preparations;
FSteps[2].ExpectedHooks[2].State := E_State.Starting;
FSteps[2].ExpectedHooks[2].Enabled := FALSE;
FSteps[2].ExpectedHooks[3].Hook := E_LifecycleHook.Tests;
FSteps[2].ExpectedHooks[3].State := E_State.Starting;
FSteps[2].ExpectedHooks[3].Enabled := FALSE;
FSteps[2].ExpectedHooks[4].Hook := E_LifecycleHook.Assertions;
FSteps[2].ExpectedHooks[4].State := E_State.Starting;
FSteps[2].ExpectedHooks[4].Enabled := FALSE;
FSteps[2].ExpectedHooks[5].Hook := E_LifecycleHook.Aggregate;
FSteps[2].ExpectedHooks[5].State := E_State.Starting;
FSteps[2].ExpectedHooks[5].Enabled := TRUE;
{endregion}

{region "03 - Wait for Preparation target"}
// Enter Preparing without evaluating Assertions; the target has not been reached.
FSteps[3].ExpectedState := E_State.Preparing;
FSteps[3].ExpectedResult := E_Result.NotEvaluated;
FSteps[3].ExpectedReady := FALSE;
FSteps[3].ExpectedPassedCount := 0;
FSteps[3].ExpectedFailedCount := 0;
FSteps[3].ExpectedHookCount := 5;
FSteps[3].ExpectedHooks[1].Hook := E_LifecycleHook.Abort;
FSteps[3].ExpectedHooks[1].State := E_State.Preparing;
FSteps[3].ExpectedHooks[1].Enabled := FALSE;
FSteps[3].ExpectedHooks[2].Hook := E_LifecycleHook.Preparations;
FSteps[3].ExpectedHooks[2].State := E_State.Preparing;
FSteps[3].ExpectedHooks[2].Enabled := TRUE;
FSteps[3].ExpectedHooks[3].Hook := E_LifecycleHook.Tests;
FSteps[3].ExpectedHooks[3].State := E_State.Preparing;
FSteps[3].ExpectedHooks[3].Enabled := FALSE;
FSteps[3].ExpectedHooks[4].Hook := E_LifecycleHook.Assertions;
FSteps[3].ExpectedHooks[4].State := E_State.Preparing;
FSteps[3].ExpectedHooks[4].Enabled := FALSE;
FSteps[3].ExpectedHooks[5].Hook := E_LifecycleHook.Aggregate;
FSteps[3].ExpectedHooks[5].State := E_State.Preparing;
FSteps[3].ExpectedHooks[5].Enabled := TRUE;
{endregion}

{region "04 - Observe target after Sequencer"}
// Publish target completion in ProcessPreparations, after this call's Sequencer has already
// run.
FSteps[4].PreparationTargetReached := TRUE;
FSteps[4].ExpectedState := E_State.Preparing;
FSteps[4].ExpectedResult := E_Result.NotEvaluated;
FSteps[4].ExpectedReady := FALSE;
FSteps[4].ExpectedPassedCount := 0;
FSteps[4].ExpectedFailedCount := 0;
FSteps[4].ExpectedHookCount := 5;
FSteps[4].ExpectedHooks[1].Hook := E_LifecycleHook.Abort;
FSteps[4].ExpectedHooks[1].State := E_State.Preparing;
FSteps[4].ExpectedHooks[1].Enabled := FALSE;
FSteps[4].ExpectedHooks[2].Hook := E_LifecycleHook.Preparations;
FSteps[4].ExpectedHooks[2].State := E_State.Preparing;
FSteps[4].ExpectedHooks[2].Enabled := TRUE;
FSteps[4].ExpectedHooks[3].Hook := E_LifecycleHook.Tests;
FSteps[4].ExpectedHooks[3].State := E_State.Preparing;
FSteps[4].ExpectedHooks[3].Enabled := FALSE;
FSteps[4].ExpectedHooks[4].Hook := E_LifecycleHook.Assertions;
FSteps[4].ExpectedHooks[4].State := E_State.Preparing;
FSteps[4].ExpectedHooks[4].Enabled := FALSE;
FSteps[4].ExpectedHooks[5].Hook := E_LifecycleHook.Aggregate;
FSteps[4].ExpectedHooks[5].State := E_State.Preparing;
FSteps[4].ExpectedHooks[5].Enabled := TRUE;
{endregion}

{region "05 - Handover to tests on next call"}
// The Sequencer consumes the previous completed observation and starts tests.
// Losing the target afterwards must not reactivate Preparation or disable test evaluation.
FSteps[5].PreparationTargetReached := FALSE;
FSteps[5].ExpectedState := E_State.Running;
FSteps[5].ExpectedResult := E_Result.NotEvaluated;
FSteps[5].ExpectedReady := FALSE;
FSteps[5].ExpectedPassedCount := 2;
FSteps[5].ExpectedFailedCount := 0;
FSteps[5].ExpectedHookCount := 5;
FSteps[5].ExpectedHooks[1].Hook := E_LifecycleHook.Abort;
FSteps[5].ExpectedHooks[1].State := E_State.Running;
FSteps[5].ExpectedHooks[1].Enabled := FALSE;
FSteps[5].ExpectedHooks[2].Hook := E_LifecycleHook.Preparations;
FSteps[5].ExpectedHooks[2].State := E_State.Running;
FSteps[5].ExpectedHooks[2].Enabled := FALSE;
FSteps[5].ExpectedHooks[3].Hook := E_LifecycleHook.Tests;
FSteps[5].ExpectedHooks[3].State := E_State.Running;
FSteps[5].ExpectedHooks[3].Enabled := TRUE;
FSteps[5].ExpectedHooks[4].Hook := E_LifecycleHook.Assertions;
FSteps[5].ExpectedHooks[4].State := E_State.Running;
FSteps[5].ExpectedHooks[4].Enabled := TRUE;
FSteps[5].ExpectedHooks[5].Hook := E_LifecycleHook.Aggregate;
FSteps[5].ExpectedHooks[5].State := E_State.Running;
FSteps[5].ExpectedHooks[5].Enabled := TRUE;
{endregion}

{region "06 - Complete inside test processing"}
// CompleteTests changes phase inside ProcessTests; subsequent Assertions must already be
// disabled.
FSteps[6].FinishTests := TRUE;
FSteps[6].ExpectedState := E_State.Completing;
FSteps[6].ExpectedResult := E_Result.Passed;
FSteps[6].ExpectedReady := FALSE;
FSteps[6].ExpectedPassedCount := 2;
FSteps[6].ExpectedFailedCount := 0;
FSteps[6].ExpectedHookCount := 5;
FSteps[6].ExpectedHooks[1].Hook := E_LifecycleHook.Abort;
FSteps[6].ExpectedHooks[1].State := E_State.Running;
FSteps[6].ExpectedHooks[1].Enabled := FALSE;
FSteps[6].ExpectedHooks[2].Hook := E_LifecycleHook.Preparations;
FSteps[6].ExpectedHooks[2].State := E_State.Running;
FSteps[6].ExpectedHooks[2].Enabled := FALSE;
FSteps[6].ExpectedHooks[3].Hook := E_LifecycleHook.Tests;
FSteps[6].ExpectedHooks[3].State := E_State.Running;
FSteps[6].ExpectedHooks[3].Enabled := TRUE;
FSteps[6].ExpectedHooks[4].Hook := E_LifecycleHook.Assertions;
FSteps[6].ExpectedHooks[4].State := E_State.Completing;
FSteps[6].ExpectedHooks[4].Enabled := FALSE;
FSteps[6].ExpectedHooks[5].Hook := E_LifecycleHook.Aggregate;
FSteps[6].ExpectedHooks[5].State := E_State.Completing;
FSteps[6].ExpectedHooks[5].Enabled := TRUE;
{endregion}

{region "07 - Observe terminal completion"}
// The following call reaches Completed; only aggregation remains in the recorded processing
// hooks.
FSteps[7].ExpectedState := E_State.Completed;
FSteps[7].ExpectedResult := E_Result.Passed;
FSteps[7].ExpectedReady := FALSE;
FSteps[7].ExpectedPassedCount := 2;
FSteps[7].ExpectedFailedCount := 0;
FSteps[7].ExpectedHookCount := 1;
FSteps[7].ExpectedHooks[1].Hook := E_LifecycleHook.Aggregate;
FSteps[7].ExpectedHooks[1].State := E_State.Completed;
FSteps[7].ExpectedHooks[1].Enabled := TRUE;
{endregion}
END_METHOD

END_FUNCTION_BLOCK

// ---- SelfTests/TestCases/TestSuite_TestCaseLifecycle/Test_LifecycleMultipleStates.TcPOU
{region 'Documentation'}
(*!
<summary>Checks two Preparation and two Test states, including immediate hook-to-hook transitions.</summary>
*)
{endregion}
FUNCTION_BLOCK Test_LifecycleMultipleStates EXTENDS TestCaseLifecycleTestBase

VAR CONSTANT
    SecondPreparationState : E_State := E_State.Preparing + 1;
    SecondTestState : E_State := E_State.Running + 1;
END_VAR

SUPER^();

{region 'Documentation'}
(*!
<summary>Defines independent per-call stimuli and expected lifecycle/hook observations.</summary>
*)
{endregion}
METHOD PROTECTED ConfigureScenario
FSubjectPreparationCount := 2;
FSubjectTestCount := 2;
FStepCount := 9;

{region "01 - Reset to Idle"}
// Establish Idle through the parent Reset request; both child results must be cleared.
FSteps[1].RequestReset := TRUE;
FSteps[1].ExpectedState := E_State.Idle;
FSteps[1].ExpectedResult := E_Result.NotEvaluated;
FSteps[1].ExpectedReady := TRUE;
FSteps[1].ExpectedPassedCount := 0;
FSteps[1].ExpectedFailedCount := 0;
FSteps[1].ExpectedHookCount := 6;
FSteps[1].ExpectedHooks[1].Hook := E_LifecycleHook.Reset;
FSteps[1].ExpectedHooks[1].State := E_State.Reset;
FSteps[1].ExpectedHooks[1].Enabled := TRUE;
FSteps[1].ExpectedHooks[2].Hook := E_LifecycleHook.Abort;
FSteps[1].ExpectedHooks[2].State := E_State.Idle;
FSteps[1].ExpectedHooks[2].Enabled := FALSE;
FSteps[1].ExpectedHooks[3].Hook := E_LifecycleHook.Preparations;
FSteps[1].ExpectedHooks[3].State := E_State.Idle;
FSteps[1].ExpectedHooks[3].Enabled := FALSE;
FSteps[1].ExpectedHooks[4].Hook := E_LifecycleHook.Tests;
FSteps[1].ExpectedHooks[4].State := E_State.Idle;
FSteps[1].ExpectedHooks[4].Enabled := FALSE;
FSteps[1].ExpectedHooks[5].Hook := E_LifecycleHook.Assertions;
FSteps[1].ExpectedHooks[5].State := E_State.Idle;
FSteps[1].ExpectedHooks[5].Enabled := FALSE;
FSteps[1].ExpectedHooks[6].Hook := E_LifecycleHook.Aggregate;
FSteps[1].ExpectedHooks[6].State := E_State.Idle;
FSteps[1].ExpectedHooks[6].Enabled := TRUE;
{endregion}

{region "02 - Accept Start"}
// Accept Start into Starting; processing and Assertion evaluation are not active yet.
FSteps[2].RequestStart := TRUE;
FSteps[2].ExpectedState := E_State.Starting;
FSteps[2].ExpectedResult := E_Result.NotEvaluated;
FSteps[2].ExpectedReady := FALSE;
FSteps[2].ExpectedPassedCount := 0;
FSteps[2].ExpectedFailedCount := 0;
FSteps[2].ExpectedHookCount := 5;
FSteps[2].ExpectedHooks[1].Hook := E_LifecycleHook.Abort;
FSteps[2].ExpectedHooks[1].State := E_State.Starting;
FSteps[2].ExpectedHooks[1].Enabled := FALSE;
FSteps[2].ExpectedHooks[2].Hook := E_LifecycleHook.Preparations;
FSteps[2].ExpectedHooks[2].State := E_State.Starting;
FSteps[2].ExpectedHooks[2].Enabled := FALSE;
FSteps[2].ExpectedHooks[3].Hook := E_LifecycleHook.Tests;
FSteps[2].ExpectedHooks[3].State := E_State.Starting;
FSteps[2].ExpectedHooks[3].Enabled := FALSE;
FSteps[2].ExpectedHooks[4].Hook := E_LifecycleHook.Assertions;
FSteps[2].ExpectedHooks[4].State := E_State.Starting;
FSteps[2].ExpectedHooks[4].Enabled := FALSE;
FSteps[2].ExpectedHooks[5].Hook := E_LifecycleHook.Aggregate;
FSteps[2].ExpectedHooks[5].State := E_State.Starting;
FSteps[2].ExpectedHooks[5].Enabled := TRUE;
{endregion}

{region "03 - Enter first Preparation state"}
// Enter Preparing without evaluating Assertions; the target has not been reached.
FSteps[3].ExpectedState := E_State.Preparing;
FSteps[3].ExpectedResult := E_Result.NotEvaluated;
FSteps[3].ExpectedReady := FALSE;
FSteps[3].ExpectedPassedCount := 0;
FSteps[3].ExpectedFailedCount := 0;
FSteps[3].ExpectedHookCount := 5;
FSteps[3].ExpectedHooks[1].Hook := E_LifecycleHook.Abort;
FSteps[3].ExpectedHooks[1].State := E_State.Preparing;
FSteps[3].ExpectedHooks[1].Enabled := FALSE;
FSteps[3].ExpectedHooks[2].Hook := E_LifecycleHook.Preparations;
FSteps[3].ExpectedHooks[2].State := E_State.Preparing;
FSteps[3].ExpectedHooks[2].Enabled := TRUE;
FSteps[3].ExpectedHooks[3].Hook := E_LifecycleHook.Tests;
FSteps[3].ExpectedHooks[3].State := E_State.Preparing;
FSteps[3].ExpectedHooks[3].Enabled := FALSE;
FSteps[3].ExpectedHooks[4].Hook := E_LifecycleHook.Assertions;
FSteps[3].ExpectedHooks[4].State := E_State.Preparing;
FSteps[3].ExpectedHooks[4].Enabled := FALSE;
FSteps[3].ExpectedHooks[5].Hook := E_LifecycleHook.Aggregate;
FSteps[3].ExpectedHooks[5].State := E_State.Preparing;
FSteps[3].ExpectedHooks[5].Enabled := TRUE;
{endregion}

{region "04 - Advance Preparation state"}
// Advance within Preparation; the entry trace records the old state, later hooks see the second
// state.
FSteps[4].AdvancePreparation := TRUE;
FSteps[4].ExpectedState := SecondPreparationState;
FSteps[4].ExpectedResult := E_Result.NotEvaluated;
FSteps[4].ExpectedReady := FALSE;
FSteps[4].ExpectedPassedCount := 0;
FSteps[4].ExpectedFailedCount := 0;
FSteps[4].ExpectedHookCount := 5;
FSteps[4].ExpectedHooks[1].Hook := E_LifecycleHook.Abort;
FSteps[4].ExpectedHooks[1].State := E_State.Preparing;
FSteps[4].ExpectedHooks[1].Enabled := FALSE;
FSteps[4].ExpectedHooks[2].Hook := E_LifecycleHook.Preparations;
FSteps[4].ExpectedHooks[2].State := E_State.Preparing;
FSteps[4].ExpectedHooks[2].Enabled := TRUE;
FSteps[4].ExpectedHooks[3].Hook := E_LifecycleHook.Tests;
FSteps[4].ExpectedHooks[3].State := SecondPreparationState;
FSteps[4].ExpectedHooks[3].Enabled := FALSE;
FSteps[4].ExpectedHooks[4].Hook := E_LifecycleHook.Assertions;
FSteps[4].ExpectedHooks[4].State := SecondPreparationState;
FSteps[4].ExpectedHooks[4].Enabled := FALSE;
FSteps[4].ExpectedHooks[5].Hook := E_LifecycleHook.Aggregate;
FSteps[4].ExpectedHooks[5].State := SecondPreparationState;
FSteps[4].ExpectedHooks[5].Enabled := TRUE;
{endregion}

{region "05 - Complete Preparation within the call"}
// Complete the reached Preparation explicitly inside its hook.
// ProcessTests and Assertions must observe Running and be enabled in this same call.
FSteps[5].FinishPreparations := TRUE;
FSteps[5].PreparationTargetReached := TRUE;
FSteps[5].ExpectedState := E_State.Running;
FSteps[5].ExpectedResult := E_Result.NotEvaluated;
FSteps[5].ExpectedReady := FALSE;
FSteps[5].ExpectedPassedCount := 2;
FSteps[5].ExpectedFailedCount := 0;
FSteps[5].ExpectedHookCount := 5;
FSteps[5].ExpectedHooks[1].Hook := E_LifecycleHook.Abort;
FSteps[5].ExpectedHooks[1].State := SecondPreparationState;
FSteps[5].ExpectedHooks[1].Enabled := FALSE;
FSteps[5].ExpectedHooks[2].Hook := E_LifecycleHook.Preparations;
FSteps[5].ExpectedHooks[2].State := SecondPreparationState;
FSteps[5].ExpectedHooks[2].Enabled := TRUE;
FSteps[5].ExpectedHooks[3].Hook := E_LifecycleHook.Tests;
FSteps[5].ExpectedHooks[3].State := E_State.Running;
FSteps[5].ExpectedHooks[3].Enabled := TRUE;
FSteps[5].ExpectedHooks[4].Hook := E_LifecycleHook.Assertions;
FSteps[5].ExpectedHooks[4].State := E_State.Running;
FSteps[5].ExpectedHooks[4].Enabled := TRUE;
FSteps[5].ExpectedHooks[5].Hook := E_LifecycleHook.Aggregate;
FSteps[5].ExpectedHooks[5].State := E_State.Running;
FSteps[5].ExpectedHooks[5].Enabled := TRUE;
{endregion}

{region "06 - Advance Test state"}
// Advance inside ProcessTests; Assertions must already observe the second Test state.
FSteps[6].AdvanceTest := TRUE;
FSteps[6].ExpectedState := SecondTestState;
FSteps[6].ExpectedResult := E_Result.NotEvaluated;
FSteps[6].ExpectedReady := FALSE;
FSteps[6].ExpectedPassedCount := 2;
FSteps[6].ExpectedFailedCount := 0;
FSteps[6].ExpectedHookCount := 5;
FSteps[6].ExpectedHooks[1].Hook := E_LifecycleHook.Abort;
FSteps[6].ExpectedHooks[1].State := E_State.Running;
FSteps[6].ExpectedHooks[1].Enabled := FALSE;
FSteps[6].ExpectedHooks[2].Hook := E_LifecycleHook.Preparations;
FSteps[6].ExpectedHooks[2].State := E_State.Running;
FSteps[6].ExpectedHooks[2].Enabled := FALSE;
FSteps[6].ExpectedHooks[3].Hook := E_LifecycleHook.Tests;
FSteps[6].ExpectedHooks[3].State := E_State.Running;
FSteps[6].ExpectedHooks[3].Enabled := TRUE;
FSteps[6].ExpectedHooks[4].Hook := E_LifecycleHook.Assertions;
FSteps[6].ExpectedHooks[4].State := SecondTestState;
FSteps[6].ExpectedHooks[4].Enabled := TRUE;
FSteps[6].ExpectedHooks[5].Hook := E_LifecycleHook.Aggregate;
FSteps[6].ExpectedHooks[5].State := SecondTestState;
FSteps[6].ExpectedHooks[5].Enabled := TRUE;
{endregion}

{region "07 - Keep second Test state active"}
// Remain in the second Test state until the concrete implementation explicitly completes it.
FSteps[7].ExpectedState := SecondTestState;
FSteps[7].ExpectedResult := E_Result.NotEvaluated;
FSteps[7].ExpectedReady := FALSE;
FSteps[7].ExpectedPassedCount := 2;
FSteps[7].ExpectedFailedCount := 0;
FSteps[7].ExpectedHookCount := 5;
FSteps[7].ExpectedHooks[1].Hook := E_LifecycleHook.Abort;
FSteps[7].ExpectedHooks[1].State := SecondTestState;
FSteps[7].ExpectedHooks[1].Enabled := FALSE;
FSteps[7].ExpectedHooks[2].Hook := E_LifecycleHook.Preparations;
FSteps[7].ExpectedHooks[2].State := SecondTestState;
FSteps[7].ExpectedHooks[2].Enabled := FALSE;
FSteps[7].ExpectedHooks[3].Hook := E_LifecycleHook.Tests;
FSteps[7].ExpectedHooks[3].State := SecondTestState;
FSteps[7].ExpectedHooks[3].Enabled := TRUE;
FSteps[7].ExpectedHooks[4].Hook := E_LifecycleHook.Assertions;
FSteps[7].ExpectedHooks[4].State := SecondTestState;
FSteps[7].ExpectedHooks[4].Enabled := TRUE;
FSteps[7].ExpectedHooks[5].Hook := E_LifecycleHook.Aggregate;
FSteps[7].ExpectedHooks[5].State := SecondTestState;
FSteps[7].ExpectedHooks[5].Enabled := TRUE;
{endregion}

{region "08 - Complete inside test processing"}
// CompleteTests changes phase inside ProcessTests; subsequent Assertions must already be
// disabled.
FSteps[8].FinishTests := TRUE;
FSteps[8].ExpectedState := E_State.Completing;
FSteps[8].ExpectedResult := E_Result.Passed;
FSteps[8].ExpectedReady := FALSE;
FSteps[8].ExpectedPassedCount := 2;
FSteps[8].ExpectedFailedCount := 0;
FSteps[8].ExpectedHookCount := 5;
FSteps[8].ExpectedHooks[1].Hook := E_LifecycleHook.Abort;
FSteps[8].ExpectedHooks[1].State := SecondTestState;
FSteps[8].ExpectedHooks[1].Enabled := FALSE;
FSteps[8].ExpectedHooks[2].Hook := E_LifecycleHook.Preparations;
FSteps[8].ExpectedHooks[2].State := SecondTestState;
FSteps[8].ExpectedHooks[2].Enabled := FALSE;
FSteps[8].ExpectedHooks[3].Hook := E_LifecycleHook.Tests;
FSteps[8].ExpectedHooks[3].State := SecondTestState;
FSteps[8].ExpectedHooks[3].Enabled := TRUE;
FSteps[8].ExpectedHooks[4].Hook := E_LifecycleHook.Assertions;
FSteps[8].ExpectedHooks[4].State := E_State.Completing;
FSteps[8].ExpectedHooks[4].Enabled := FALSE;
FSteps[8].ExpectedHooks[5].Hook := E_LifecycleHook.Aggregate;
FSteps[8].ExpectedHooks[5].State := E_State.Completing;
FSteps[8].ExpectedHooks[5].Enabled := TRUE;
{endregion}

{region "09 - Observe terminal completion"}
// The following call reaches Completed; only aggregation remains in the recorded processing
// hooks.
FSteps[9].ExpectedState := E_State.Completed;
FSteps[9].ExpectedResult := E_Result.Passed;
FSteps[9].ExpectedReady := FALSE;
FSteps[9].ExpectedPassedCount := 2;
FSteps[9].ExpectedFailedCount := 0;
FSteps[9].ExpectedHookCount := 1;
FSteps[9].ExpectedHooks[1].Hook := E_LifecycleHook.Aggregate;
FSteps[9].ExpectedHooks[1].State := E_State.Completed;
FSteps[9].ExpectedHooks[1].Enabled := TRUE;
{endregion}
END_METHOD

END_FUNCTION_BLOCK

// ---- SelfTests/TestCases/TestSuite_TestCaseLifecycle/Test_LifecycleAlreadyPrepared.TcPOU
{region 'Documentation'}
(*!
<summary>Checks that an already reached target skips active Preparation without suppressing Test execution.</summary>
*)
{endregion}
FUNCTION_BLOCK Test_LifecycleAlreadyPrepared EXTENDS TestCaseLifecycleTestBase

SUPER^();

{region 'Documentation'}
(*!
<summary>Defines independent per-call stimuli and expected lifecycle/hook observations.</summary>
*)
{endregion}
METHOD PROTECTED ConfigureScenario
FSubjectPreparationCount := 1;
FSubjectTestCount := 1;
FStepCount := 6;

{region "01 - Reset to Idle"}
// Establish Idle through the parent Reset request; both child results must be cleared.
FSteps[1].RequestReset := TRUE;
FSteps[1].ExpectedState := E_State.Idle;
FSteps[1].ExpectedResult := E_Result.NotEvaluated;
FSteps[1].ExpectedReady := TRUE;
FSteps[1].ExpectedPassedCount := 0;
FSteps[1].ExpectedFailedCount := 0;
FSteps[1].ExpectedHookCount := 6;
FSteps[1].ExpectedHooks[1].Hook := E_LifecycleHook.Reset;
FSteps[1].ExpectedHooks[1].State := E_State.Reset;
FSteps[1].ExpectedHooks[1].Enabled := TRUE;
FSteps[1].ExpectedHooks[2].Hook := E_LifecycleHook.Abort;
FSteps[1].ExpectedHooks[2].State := E_State.Idle;
FSteps[1].ExpectedHooks[2].Enabled := FALSE;
FSteps[1].ExpectedHooks[3].Hook := E_LifecycleHook.Preparations;
FSteps[1].ExpectedHooks[3].State := E_State.Idle;
FSteps[1].ExpectedHooks[3].Enabled := FALSE;
FSteps[1].ExpectedHooks[4].Hook := E_LifecycleHook.Tests;
FSteps[1].ExpectedHooks[4].State := E_State.Idle;
FSteps[1].ExpectedHooks[4].Enabled := FALSE;
FSteps[1].ExpectedHooks[5].Hook := E_LifecycleHook.Assertions;
FSteps[1].ExpectedHooks[5].State := E_State.Idle;
FSteps[1].ExpectedHooks[5].Enabled := FALSE;
FSteps[1].ExpectedHooks[6].Hook := E_LifecycleHook.Aggregate;
FSteps[1].ExpectedHooks[6].State := E_State.Idle;
FSteps[1].ExpectedHooks[6].Enabled := TRUE;
{endregion}

{region "02 - Observe target before Start"}
// Observe the reached target while Idle, before requesting execution.
FSteps[2].PreparationTargetReached := TRUE;
FSteps[2].ExpectedState := E_State.Idle;
FSteps[2].ExpectedResult := E_Result.NotEvaluated;
FSteps[2].ExpectedReady := TRUE;
FSteps[2].ExpectedPassedCount := 0;
FSteps[2].ExpectedFailedCount := 0;
FSteps[2].ExpectedHookCount := 5;
FSteps[2].ExpectedHooks[1].Hook := E_LifecycleHook.Abort;
FSteps[2].ExpectedHooks[1].State := E_State.Idle;
FSteps[2].ExpectedHooks[1].Enabled := FALSE;
FSteps[2].ExpectedHooks[2].Hook := E_LifecycleHook.Preparations;
FSteps[2].ExpectedHooks[2].State := E_State.Idle;
FSteps[2].ExpectedHooks[2].Enabled := FALSE;
FSteps[2].ExpectedHooks[3].Hook := E_LifecycleHook.Tests;
FSteps[2].ExpectedHooks[3].State := E_State.Idle;
FSteps[2].ExpectedHooks[3].Enabled := FALSE;
FSteps[2].ExpectedHooks[4].Hook := E_LifecycleHook.Assertions;
FSteps[2].ExpectedHooks[4].State := E_State.Idle;
FSteps[2].ExpectedHooks[4].Enabled := FALSE;
FSteps[2].ExpectedHooks[5].Hook := E_LifecycleHook.Aggregate;
FSteps[2].ExpectedHooks[5].State := E_State.Idle;
FSteps[2].ExpectedHooks[5].Enabled := TRUE;
{endregion}

{region "03 - Start with completed Preparation"}
// Start with a completed Preparation observation already available.
FSteps[3].RequestStart := TRUE;
FSteps[3].PreparationTargetReached := TRUE;
FSteps[3].ExpectedState := E_State.Starting;
FSteps[3].ExpectedResult := E_Result.NotEvaluated;
FSteps[3].ExpectedReady := FALSE;
FSteps[3].ExpectedPassedCount := 0;
FSteps[3].ExpectedFailedCount := 0;
FSteps[3].ExpectedHookCount := 5;
FSteps[3].ExpectedHooks[1].Hook := E_LifecycleHook.Abort;
FSteps[3].ExpectedHooks[1].State := E_State.Starting;
FSteps[3].ExpectedHooks[1].Enabled := FALSE;
FSteps[3].ExpectedHooks[2].Hook := E_LifecycleHook.Preparations;
FSteps[3].ExpectedHooks[2].State := E_State.Starting;
FSteps[3].ExpectedHooks[2].Enabled := FALSE;
FSteps[3].ExpectedHooks[3].Hook := E_LifecycleHook.Tests;
FSteps[3].ExpectedHooks[3].State := E_State.Starting;
FSteps[3].ExpectedHooks[3].Enabled := FALSE;
FSteps[3].ExpectedHooks[4].Hook := E_LifecycleHook.Assertions;
FSteps[3].ExpectedHooks[4].State := E_State.Starting;
FSteps[3].ExpectedHooks[4].Enabled := FALSE;
FSteps[3].ExpectedHooks[5].Hook := E_LifecycleHook.Aggregate;
FSteps[3].ExpectedHooks[5].State := E_State.Starting;
FSteps[3].ExpectedHooks[5].Enabled := TRUE;
{endregion}

{region "04 - Skip active Preparation"}
// Skip active Preparation based on the previous observation.
// The current target may disappear during testing without blocking Running.
FSteps[4].PreparationTargetReached := FALSE;
FSteps[4].ExpectedState := E_State.Running;
FSteps[4].ExpectedResult := E_Result.NotEvaluated;
FSteps[4].ExpectedReady := FALSE;
FSteps[4].ExpectedPassedCount := 2;
FSteps[4].ExpectedFailedCount := 0;
FSteps[4].ExpectedHookCount := 5;
FSteps[4].ExpectedHooks[1].Hook := E_LifecycleHook.Abort;
FSteps[4].ExpectedHooks[1].State := E_State.Running;
FSteps[4].ExpectedHooks[1].Enabled := FALSE;
FSteps[4].ExpectedHooks[2].Hook := E_LifecycleHook.Preparations;
FSteps[4].ExpectedHooks[2].State := E_State.Running;
FSteps[4].ExpectedHooks[2].Enabled := FALSE;
FSteps[4].ExpectedHooks[3].Hook := E_LifecycleHook.Tests;
FSteps[4].ExpectedHooks[3].State := E_State.Running;
FSteps[4].ExpectedHooks[3].Enabled := TRUE;
FSteps[4].ExpectedHooks[4].Hook := E_LifecycleHook.Assertions;
FSteps[4].ExpectedHooks[4].State := E_State.Running;
FSteps[4].ExpectedHooks[4].Enabled := TRUE;
FSteps[4].ExpectedHooks[5].Hook := E_LifecycleHook.Aggregate;
FSteps[4].ExpectedHooks[5].State := E_State.Running;
FSteps[4].ExpectedHooks[5].Enabled := TRUE;
{endregion}

{region "05 - Complete inside test processing"}
// CompleteTests changes phase inside ProcessTests; subsequent Assertions must already be
// disabled.
FSteps[5].FinishTests := TRUE;
FSteps[5].ExpectedState := E_State.Completing;
FSteps[5].ExpectedResult := E_Result.Passed;
FSteps[5].ExpectedReady := FALSE;
FSteps[5].ExpectedPassedCount := 2;
FSteps[5].ExpectedFailedCount := 0;
FSteps[5].ExpectedHookCount := 5;
FSteps[5].ExpectedHooks[1].Hook := E_LifecycleHook.Abort;
FSteps[5].ExpectedHooks[1].State := E_State.Running;
FSteps[5].ExpectedHooks[1].Enabled := FALSE;
FSteps[5].ExpectedHooks[2].Hook := E_LifecycleHook.Preparations;
FSteps[5].ExpectedHooks[2].State := E_State.Running;
FSteps[5].ExpectedHooks[2].Enabled := FALSE;
FSteps[5].ExpectedHooks[3].Hook := E_LifecycleHook.Tests;
FSteps[5].ExpectedHooks[3].State := E_State.Running;
FSteps[5].ExpectedHooks[3].Enabled := TRUE;
FSteps[5].ExpectedHooks[4].Hook := E_LifecycleHook.Assertions;
FSteps[5].ExpectedHooks[4].State := E_State.Completing;
FSteps[5].ExpectedHooks[4].Enabled := FALSE;
FSteps[5].ExpectedHooks[5].Hook := E_LifecycleHook.Aggregate;
FSteps[5].ExpectedHooks[5].State := E_State.Completing;
FSteps[5].ExpectedHooks[5].Enabled := TRUE;
{endregion}

{region "06 - Observe terminal completion"}
// The following call reaches Completed; only aggregation remains in the recorded processing
// hooks.
FSteps[6].ExpectedState := E_State.Completed;
FSteps[6].ExpectedResult := E_Result.Passed;
FSteps[6].ExpectedReady := FALSE;
FSteps[6].ExpectedPassedCount := 2;
FSteps[6].ExpectedFailedCount := 0;
FSteps[6].ExpectedHookCount := 1;
FSteps[6].ExpectedHooks[1].Hook := E_LifecycleHook.Aggregate;
FSteps[6].ExpectedHooks[1].State := E_State.Completed;
FSteps[6].ExpectedHooks[1].Enabled := TRUE;
{endregion}
END_METHOD

END_FUNCTION_BLOCK

// ---- SelfTests/TestCases/TestSuite_TestCaseLifecycle/Test_LifecycleFailedResult.TcPOU
{region 'Documentation'}
(*!
<summary>
Checks mixed Assertion aggregation, continued execution after Failed and explicit Failed finalization.
</summary>
*)
{endregion}
FUNCTION_BLOCK Test_LifecycleFailedResult EXTENDS TestCaseLifecycleTestBase

SUPER^();

{region 'Documentation'}
(*!
<summary>Defines an independent cycle trace including mixed Passed/Failed results.</summary>
*)
{endregion}
METHOD PROTECTED ConfigureScenario
FSubjectPreparationCount := 0;
FSubjectTestCount := 1;
FStepCount := 6;

{region "01 - Reset to Idle"}
// Establish Idle through the parent Reset request; both child results must be cleared.
FSteps[1].RequestReset := TRUE;
FSteps[1].ExpectedState := E_State.Idle;
FSteps[1].ExpectedResult := E_Result.NotEvaluated;
FSteps[1].ExpectedReady := TRUE;
FSteps[1].ExpectedPassedCount := 0;
FSteps[1].ExpectedFailedCount := 0;
FSteps[1].ExpectedHookCount := 6;
FSteps[1].ExpectedHooks[1].Hook := E_LifecycleHook.Reset;
FSteps[1].ExpectedHooks[1].State := E_State.Reset;
FSteps[1].ExpectedHooks[1].Enabled := TRUE;
FSteps[1].ExpectedHooks[2].Hook := E_LifecycleHook.Abort;
FSteps[1].ExpectedHooks[2].State := E_State.Idle;
FSteps[1].ExpectedHooks[2].Enabled := FALSE;
FSteps[1].ExpectedHooks[3].Hook := E_LifecycleHook.Preparations;
FSteps[1].ExpectedHooks[3].State := E_State.Idle;
FSteps[1].ExpectedHooks[3].Enabled := FALSE;
FSteps[1].ExpectedHooks[4].Hook := E_LifecycleHook.Tests;
FSteps[1].ExpectedHooks[4].State := E_State.Idle;
FSteps[1].ExpectedHooks[4].Enabled := FALSE;
FSteps[1].ExpectedHooks[5].Hook := E_LifecycleHook.Assertions;
FSteps[1].ExpectedHooks[5].State := E_State.Idle;
FSteps[1].ExpectedHooks[5].Enabled := FALSE;
FSteps[1].ExpectedHooks[6].Hook := E_LifecycleHook.Aggregate;
FSteps[1].ExpectedHooks[6].State := E_State.Idle;
FSteps[1].ExpectedHooks[6].Enabled := TRUE;
{endregion}

{region "02 - Accept Start"}
// Accept Start into Starting; processing and Assertion evaluation are not active yet.
FSteps[2].RequestStart := TRUE;
FSteps[2].ExpectedState := E_State.Starting;
FSteps[2].ExpectedResult := E_Result.NotEvaluated;
FSteps[2].ExpectedReady := FALSE;
FSteps[2].ExpectedPassedCount := 0;
FSteps[2].ExpectedFailedCount := 0;
FSteps[2].ExpectedHookCount := 5;
FSteps[2].ExpectedHooks[1].Hook := E_LifecycleHook.Abort;
FSteps[2].ExpectedHooks[1].State := E_State.Starting;
FSteps[2].ExpectedHooks[1].Enabled := FALSE;
FSteps[2].ExpectedHooks[2].Hook := E_LifecycleHook.Preparations;
FSteps[2].ExpectedHooks[2].State := E_State.Starting;
FSteps[2].ExpectedHooks[2].Enabled := FALSE;
FSteps[2].ExpectedHooks[3].Hook := E_LifecycleHook.Tests;
FSteps[2].ExpectedHooks[3].State := E_State.Starting;
FSteps[2].ExpectedHooks[3].Enabled := FALSE;
FSteps[2].ExpectedHooks[4].Hook := E_LifecycleHook.Assertions;
FSteps[2].ExpectedHooks[4].State := E_State.Starting;
FSteps[2].ExpectedHooks[4].Enabled := FALSE;
FSteps[2].ExpectedHooks[5].Hook := E_LifecycleHook.Aggregate;
FSteps[2].ExpectedHooks[5].State := E_State.Starting;
FSteps[2].ExpectedHooks[5].Enabled := TRUE;
{endregion}

{region "03 - Generate one child failure"}
// Make Condition fail while ReferenceCondition passes; counters expose both outcomes during
// Running.
FSteps[3].AssertionCondition := FALSE;
FSteps[3].ExpectedState := E_State.Running;
FSteps[3].ExpectedResult := E_Result.NotEvaluated;
FSteps[3].ExpectedReady := FALSE;
FSteps[3].ExpectedPassedCount := 1;
FSteps[3].ExpectedFailedCount := 1;
FSteps[3].ExpectedHookCount := 5;
FSteps[3].ExpectedHooks[1].Hook := E_LifecycleHook.Abort;
FSteps[3].ExpectedHooks[1].State := E_State.Running;
FSteps[3].ExpectedHooks[1].Enabled := FALSE;
FSteps[3].ExpectedHooks[2].Hook := E_LifecycleHook.Preparations;
FSteps[3].ExpectedHooks[2].State := E_State.Running;
FSteps[3].ExpectedHooks[2].Enabled := FALSE;
FSteps[3].ExpectedHooks[3].Hook := E_LifecycleHook.Tests;
FSteps[3].ExpectedHooks[3].State := E_State.Running;
FSteps[3].ExpectedHooks[3].Enabled := TRUE;
FSteps[3].ExpectedHooks[4].Hook := E_LifecycleHook.Assertions;
FSteps[3].ExpectedHooks[4].State := E_State.Running;
FSteps[3].ExpectedHooks[4].Enabled := TRUE;
FSteps[3].ExpectedHooks[5].Hook := E_LifecycleHook.Aggregate;
FSteps[3].ExpectedHooks[5].State := E_State.Running;
FSteps[3].ExpectedHooks[5].Enabled := TRUE;
{endregion}

{region "04 - Preserve latched failure"}
// Restore Condition input to TRUE; the already latched Failed result must not recover without
// Reset.
FSteps[4].ExpectedState := E_State.Running;
FSteps[4].ExpectedResult := E_Result.NotEvaluated;
FSteps[4].ExpectedReady := FALSE;
FSteps[4].ExpectedPassedCount := 1;
FSteps[4].ExpectedFailedCount := 1;
FSteps[4].ExpectedHookCount := 5;
FSteps[4].ExpectedHooks[1].Hook := E_LifecycleHook.Abort;
FSteps[4].ExpectedHooks[1].State := E_State.Running;
FSteps[4].ExpectedHooks[1].Enabled := FALSE;
FSteps[4].ExpectedHooks[2].Hook := E_LifecycleHook.Preparations;
FSteps[4].ExpectedHooks[2].State := E_State.Running;
FSteps[4].ExpectedHooks[2].Enabled := FALSE;
FSteps[4].ExpectedHooks[3].Hook := E_LifecycleHook.Tests;
FSteps[4].ExpectedHooks[3].State := E_State.Running;
FSteps[4].ExpectedHooks[3].Enabled := TRUE;
FSteps[4].ExpectedHooks[4].Hook := E_LifecycleHook.Assertions;
FSteps[4].ExpectedHooks[4].State := E_State.Running;
FSteps[4].ExpectedHooks[4].Enabled := TRUE;
FSteps[4].ExpectedHooks[5].Hook := E_LifecycleHook.Aggregate;
FSteps[4].ExpectedHooks[5].State := E_State.Running;
FSteps[4].ExpectedHooks[5].Enabled := TRUE;
{endregion}

{region "05 - Finalize with Failed"}
// Complete execution; the held child failure must now become the Test Case's Failed result.
FSteps[5].FinishTests := TRUE;
FSteps[5].ExpectedState := E_State.Completing;
FSteps[5].ExpectedResult := E_Result.Failed;
FSteps[5].ExpectedReady := FALSE;
FSteps[5].ExpectedPassedCount := 1;
FSteps[5].ExpectedFailedCount := 1;
FSteps[5].ExpectedHookCount := 5;
FSteps[5].ExpectedHooks[1].Hook := E_LifecycleHook.Abort;
FSteps[5].ExpectedHooks[1].State := E_State.Running;
FSteps[5].ExpectedHooks[1].Enabled := FALSE;
FSteps[5].ExpectedHooks[2].Hook := E_LifecycleHook.Preparations;
FSteps[5].ExpectedHooks[2].State := E_State.Running;
FSteps[5].ExpectedHooks[2].Enabled := FALSE;
FSteps[5].ExpectedHooks[3].Hook := E_LifecycleHook.Tests;
FSteps[5].ExpectedHooks[3].State := E_State.Running;
FSteps[5].ExpectedHooks[3].Enabled := TRUE;
FSteps[5].ExpectedHooks[4].Hook := E_LifecycleHook.Assertions;
FSteps[5].ExpectedHooks[4].State := E_State.Completing;
FSteps[5].ExpectedHooks[4].Enabled := FALSE;
FSteps[5].ExpectedHooks[5].Hook := E_LifecycleHook.Aggregate;
FSteps[5].ExpectedHooks[5].State := E_State.Completing;
FSteps[5].ExpectedHooks[5].Enabled := TRUE;
{endregion}

{region "06 - Observe terminal completion"}
// The following call reaches Completed; only aggregation remains in the recorded processing
// hooks.
FSteps[6].ExpectedState := E_State.Completed;
FSteps[6].ExpectedResult := E_Result.Failed;
FSteps[6].ExpectedReady := FALSE;
FSteps[6].ExpectedPassedCount := 1;
FSteps[6].ExpectedFailedCount := 1;
FSteps[6].ExpectedHookCount := 1;
FSteps[6].ExpectedHooks[1].Hook := E_LifecycleHook.Aggregate;
FSteps[6].ExpectedHooks[1].State := E_State.Completed;
FSteps[6].ExpectedHooks[1].Enabled := TRUE;
{endregion}
END_METHOD

END_FUNCTION_BLOCK

// ---- SelfTests/TestCases/TestSuite_TestCaseLifecycle/Test_LifecycleAbort.TcPOU
{region 'Documentation'}
(*!
<summary>Checks held Abort cleanup and explicit completion without further enabled test work.</summary>
*)
{endregion}
FUNCTION_BLOCK Test_LifecycleAbort EXTENDS TestCaseLifecycleTestBase

SUPER^();

{region 'Documentation'}
(*!
<summary>Defines explicit exceptional-path stimuli and contract-derived observations.</summary>
*)
{endregion}
METHOD PROTECTED ConfigureScenario
FSubjectPreparationCount := 0;
FSubjectTestCount := 1;
FStepCount := 7;

{region "01 - Reset to Idle"}
// Establish Idle through the parent Reset request; both child results must be cleared.
FSteps[1].RequestReset := TRUE;
FSteps[1].ExpectedState := E_State.Idle;
FSteps[1].ExpectedResult := E_Result.NotEvaluated;
FSteps[1].ExpectedReady := TRUE;
FSteps[1].ExpectedPassedCount := 0;
FSteps[1].ExpectedFailedCount := 0;
FSteps[1].ExpectedHookCount := 6;
FSteps[1].ExpectedHooks[1].Hook := E_LifecycleHook.Reset;
FSteps[1].ExpectedHooks[1].State := E_State.Reset;
FSteps[1].ExpectedHooks[1].Enabled := TRUE;
FSteps[1].ExpectedHooks[2].Hook := E_LifecycleHook.Abort;
FSteps[1].ExpectedHooks[2].State := E_State.Idle;
FSteps[1].ExpectedHooks[2].Enabled := FALSE;
FSteps[1].ExpectedHooks[3].Hook := E_LifecycleHook.Preparations;
FSteps[1].ExpectedHooks[3].State := E_State.Idle;
FSteps[1].ExpectedHooks[3].Enabled := FALSE;
FSteps[1].ExpectedHooks[4].Hook := E_LifecycleHook.Tests;
FSteps[1].ExpectedHooks[4].State := E_State.Idle;
FSteps[1].ExpectedHooks[4].Enabled := FALSE;
FSteps[1].ExpectedHooks[5].Hook := E_LifecycleHook.Assertions;
FSteps[1].ExpectedHooks[5].State := E_State.Idle;
FSteps[1].ExpectedHooks[5].Enabled := FALSE;
FSteps[1].ExpectedHooks[6].Hook := E_LifecycleHook.Aggregate;
FSteps[1].ExpectedHooks[6].State := E_State.Idle;
FSteps[1].ExpectedHooks[6].Enabled := TRUE;
{endregion}

{region "02 - Accept Start"}
// Accept Start into Starting; processing and Assertion evaluation are not active yet.
FSteps[2].RequestStart := TRUE;
FSteps[2].ExpectedState := E_State.Starting;
FSteps[2].ExpectedResult := E_Result.NotEvaluated;
FSteps[2].ExpectedReady := FALSE;
FSteps[2].ExpectedPassedCount := 0;
FSteps[2].ExpectedFailedCount := 0;
FSteps[2].ExpectedHookCount := 5;
FSteps[2].ExpectedHooks[1].Hook := E_LifecycleHook.Abort;
FSteps[2].ExpectedHooks[1].State := E_State.Starting;
FSteps[2].ExpectedHooks[1].Enabled := FALSE;
FSteps[2].ExpectedHooks[2].Hook := E_LifecycleHook.Preparations;
FSteps[2].ExpectedHooks[2].State := E_State.Starting;
FSteps[2].ExpectedHooks[2].Enabled := FALSE;
FSteps[2].ExpectedHooks[3].Hook := E_LifecycleHook.Tests;
FSteps[2].ExpectedHooks[3].State := E_State.Starting;
FSteps[2].ExpectedHooks[3].Enabled := FALSE;
FSteps[2].ExpectedHooks[4].Hook := E_LifecycleHook.Assertions;
FSteps[2].ExpectedHooks[4].State := E_State.Starting;
FSteps[2].ExpectedHooks[4].Enabled := FALSE;
FSteps[2].ExpectedHooks[5].Hook := E_LifecycleHook.Aggregate;
FSteps[2].ExpectedHooks[5].State := E_State.Starting;
FSteps[2].ExpectedHooks[5].Enabled := TRUE;
{endregion}

{region "03 - Establish active execution"}
// Enter Running and evaluate both children; owner Result stays NotEvaluated until finalization.
FSteps[3].ExpectedState := E_State.Running;
FSteps[3].ExpectedResult := E_Result.NotEvaluated;
FSteps[3].ExpectedReady := FALSE;
FSteps[3].ExpectedPassedCount := 2;
FSteps[3].ExpectedFailedCount := 0;
FSteps[3].ExpectedHookCount := 5;
FSteps[3].ExpectedHooks[1].Hook := E_LifecycleHook.Abort;
FSteps[3].ExpectedHooks[1].State := E_State.Running;
FSteps[3].ExpectedHooks[1].Enabled := FALSE;
FSteps[3].ExpectedHooks[2].Hook := E_LifecycleHook.Preparations;
FSteps[3].ExpectedHooks[2].State := E_State.Running;
FSteps[3].ExpectedHooks[2].Enabled := FALSE;
FSteps[3].ExpectedHooks[3].Hook := E_LifecycleHook.Tests;
FSteps[3].ExpectedHooks[3].State := E_State.Running;
FSteps[3].ExpectedHooks[3].Enabled := TRUE;
FSteps[3].ExpectedHooks[4].Hook := E_LifecycleHook.Assertions;
FSteps[3].ExpectedHooks[4].State := E_State.Running;
FSteps[3].ExpectedHooks[4].Enabled := TRUE;
FSteps[3].ExpectedHooks[5].Hook := E_LifecycleHook.Aggregate;
FSteps[3].ExpectedHooks[5].State := E_State.Running;
FSteps[3].ExpectedHooks[5].Enabled := TRUE;
{endregion}

{region "04 - Request Abort and hold cleanup"}
// Request Abort and withhold cleanup completion; retain child results while entering Aborting.
FSteps[4].RequestAbort := TRUE;
FSteps[4].AbortCompleted := FALSE;
FSteps[4].ExpectedState := E_State.Aborting;
FSteps[4].ExpectedResult := E_Result.Abort;
FSteps[4].ExpectedReady := FALSE;
FSteps[4].ExpectedPassedCount := 2;
FSteps[4].ExpectedFailedCount := 0;
FSteps[4].ExpectedHookCount := 5;
FSteps[4].ExpectedHooks[1].Hook := E_LifecycleHook.Abort;
FSteps[4].ExpectedHooks[1].State := E_State.Aborting;
FSteps[4].ExpectedHooks[1].Enabled := TRUE;
FSteps[4].ExpectedHooks[2].Hook := E_LifecycleHook.Preparations;
FSteps[4].ExpectedHooks[2].State := E_State.Aborting;
FSteps[4].ExpectedHooks[2].Enabled := FALSE;
FSteps[4].ExpectedHooks[3].Hook := E_LifecycleHook.Tests;
FSteps[4].ExpectedHooks[3].State := E_State.Aborting;
FSteps[4].ExpectedHooks[3].Enabled := FALSE;
FSteps[4].ExpectedHooks[4].Hook := E_LifecycleHook.Assertions;
FSteps[4].ExpectedHooks[4].State := E_State.Aborting;
FSteps[4].ExpectedHooks[4].Enabled := FALSE;
FSteps[4].ExpectedHooks[5].Hook := E_LifecycleHook.Aggregate;
FSteps[4].ExpectedHooks[5].State := E_State.Aborting;
FSteps[4].ExpectedHooks[5].Enabled := TRUE;
{endregion}

{region "05 - Continue pending cleanup"}
// Continue active cleanup without a second Abort request; do not finalize before
// acknowledgement.
FSteps[5].AbortCompleted := FALSE;
FSteps[5].ExpectedState := E_State.Aborting;
FSteps[5].ExpectedResult := E_Result.Abort;
FSteps[5].ExpectedReady := FALSE;
FSteps[5].ExpectedPassedCount := 2;
FSteps[5].ExpectedFailedCount := 0;
FSteps[5].ExpectedHookCount := 5;
FSteps[5].ExpectedHooks[1].Hook := E_LifecycleHook.Abort;
FSteps[5].ExpectedHooks[1].State := E_State.Aborting;
FSteps[5].ExpectedHooks[1].Enabled := TRUE;
FSteps[5].ExpectedHooks[2].Hook := E_LifecycleHook.Preparations;
FSteps[5].ExpectedHooks[2].State := E_State.Aborting;
FSteps[5].ExpectedHooks[2].Enabled := FALSE;
FSteps[5].ExpectedHooks[3].Hook := E_LifecycleHook.Tests;
FSteps[5].ExpectedHooks[3].State := E_State.Aborting;
FSteps[5].ExpectedHooks[3].Enabled := FALSE;
FSteps[5].ExpectedHooks[4].Hook := E_LifecycleHook.Assertions;
FSteps[5].ExpectedHooks[4].State := E_State.Aborting;
FSteps[5].ExpectedHooks[4].Enabled := FALSE;
FSteps[5].ExpectedHooks[5].Hook := E_LifecycleHook.Aggregate;
FSteps[5].ExpectedHooks[5].State := E_State.Aborting;
FSteps[5].ExpectedHooks[5].Enabled := TRUE;
{endregion}

{region "06 - Acknowledge Abort cleanup"}
// Release AbortCompleted through its default TRUE value.
// The Abort hook enters Aborting, then all following hooks observe Completing.
FSteps[6].ExpectedState := E_State.Completing;
FSteps[6].ExpectedResult := E_Result.Abort;
FSteps[6].ExpectedReady := FALSE;
FSteps[6].ExpectedPassedCount := 2;
FSteps[6].ExpectedFailedCount := 0;
FSteps[6].ExpectedHookCount := 5;
FSteps[6].ExpectedHooks[1].Hook := E_LifecycleHook.Abort;
FSteps[6].ExpectedHooks[1].State := E_State.Aborting;
FSteps[6].ExpectedHooks[1].Enabled := TRUE;
FSteps[6].ExpectedHooks[2].Hook := E_LifecycleHook.Preparations;
FSteps[6].ExpectedHooks[2].State := E_State.Completing;
FSteps[6].ExpectedHooks[2].Enabled := FALSE;
FSteps[6].ExpectedHooks[3].Hook := E_LifecycleHook.Tests;
FSteps[6].ExpectedHooks[3].State := E_State.Completing;
FSteps[6].ExpectedHooks[3].Enabled := FALSE;
FSteps[6].ExpectedHooks[4].Hook := E_LifecycleHook.Assertions;
FSteps[6].ExpectedHooks[4].State := E_State.Completing;
FSteps[6].ExpectedHooks[4].Enabled := FALSE;
FSteps[6].ExpectedHooks[5].Hook := E_LifecycleHook.Aggregate;
FSteps[6].ExpectedHooks[5].State := E_State.Completing;
FSteps[6].ExpectedHooks[5].Enabled := TRUE;
{endregion}

{region "07 - Observe terminal Abort"}
// The following call reaches Completed; only aggregation remains in the recorded processing
// hooks.
FSteps[7].ExpectedState := E_State.Completed;
FSteps[7].ExpectedResult := E_Result.Abort;
FSteps[7].ExpectedReady := FALSE;
FSteps[7].ExpectedPassedCount := 2;
FSteps[7].ExpectedFailedCount := 0;
FSteps[7].ExpectedHookCount := 1;
FSteps[7].ExpectedHooks[1].Hook := E_LifecycleHook.Aggregate;
FSteps[7].ExpectedHooks[1].State := E_State.Completed;
FSteps[7].ExpectedHooks[1].Enabled := TRUE;
{endregion}
END_METHOD

END_FUNCTION_BLOCK

// ---- SelfTests/TestCases/TestSuite_TestCaseLifecycle/Test_LifecycleAbortError.TcPOU
{region 'Documentation'}
(*!
<summary>Checks escalation from Abort to Error while cleanup is still pending.</summary>
*)
{endregion}
FUNCTION_BLOCK Test_LifecycleAbortError EXTENDS TestCaseLifecycleTestBase

SUPER^();

{region 'Documentation'}
(*!
<summary>Defines explicit exceptional-path stimuli and contract-derived observations.</summary>
*)
{endregion}
METHOD PROTECTED ConfigureScenario
FSubjectPreparationCount := 0;
FSubjectTestCount := 1;
FStepCount := 7;

{region "01 - Reset to Idle"}
// Establish Idle through the parent Reset request; both child results must be cleared.
FSteps[1].RequestReset := TRUE;
FSteps[1].ExpectedState := E_State.Idle;
FSteps[1].ExpectedResult := E_Result.NotEvaluated;
FSteps[1].ExpectedReady := TRUE;
FSteps[1].ExpectedPassedCount := 0;
FSteps[1].ExpectedFailedCount := 0;
FSteps[1].ExpectedHookCount := 6;
FSteps[1].ExpectedHooks[1].Hook := E_LifecycleHook.Reset;
FSteps[1].ExpectedHooks[1].State := E_State.Reset;
FSteps[1].ExpectedHooks[1].Enabled := TRUE;
FSteps[1].ExpectedHooks[2].Hook := E_LifecycleHook.Abort;
FSteps[1].ExpectedHooks[2].State := E_State.Idle;
FSteps[1].ExpectedHooks[2].Enabled := FALSE;
FSteps[1].ExpectedHooks[3].Hook := E_LifecycleHook.Preparations;
FSteps[1].ExpectedHooks[3].State := E_State.Idle;
FSteps[1].ExpectedHooks[3].Enabled := FALSE;
FSteps[1].ExpectedHooks[4].Hook := E_LifecycleHook.Tests;
FSteps[1].ExpectedHooks[4].State := E_State.Idle;
FSteps[1].ExpectedHooks[4].Enabled := FALSE;
FSteps[1].ExpectedHooks[5].Hook := E_LifecycleHook.Assertions;
FSteps[1].ExpectedHooks[5].State := E_State.Idle;
FSteps[1].ExpectedHooks[5].Enabled := FALSE;
FSteps[1].ExpectedHooks[6].Hook := E_LifecycleHook.Aggregate;
FSteps[1].ExpectedHooks[6].State := E_State.Idle;
FSteps[1].ExpectedHooks[6].Enabled := TRUE;
{endregion}

{region "02 - Accept Start"}
// Accept Start into Starting; processing and Assertion evaluation are not active yet.
FSteps[2].RequestStart := TRUE;
FSteps[2].ExpectedState := E_State.Starting;
FSteps[2].ExpectedResult := E_Result.NotEvaluated;
FSteps[2].ExpectedReady := FALSE;
FSteps[2].ExpectedPassedCount := 0;
FSteps[2].ExpectedFailedCount := 0;
FSteps[2].ExpectedHookCount := 5;
FSteps[2].ExpectedHooks[1].Hook := E_LifecycleHook.Abort;
FSteps[2].ExpectedHooks[1].State := E_State.Starting;
FSteps[2].ExpectedHooks[1].Enabled := FALSE;
FSteps[2].ExpectedHooks[2].Hook := E_LifecycleHook.Preparations;
FSteps[2].ExpectedHooks[2].State := E_State.Starting;
FSteps[2].ExpectedHooks[2].Enabled := FALSE;
FSteps[2].ExpectedHooks[3].Hook := E_LifecycleHook.Tests;
FSteps[2].ExpectedHooks[3].State := E_State.Starting;
FSteps[2].ExpectedHooks[3].Enabled := FALSE;
FSteps[2].ExpectedHooks[4].Hook := E_LifecycleHook.Assertions;
FSteps[2].ExpectedHooks[4].State := E_State.Starting;
FSteps[2].ExpectedHooks[4].Enabled := FALSE;
FSteps[2].ExpectedHooks[5].Hook := E_LifecycleHook.Aggregate;
FSteps[2].ExpectedHooks[5].State := E_State.Starting;
FSteps[2].ExpectedHooks[5].Enabled := TRUE;
{endregion}

{region "03 - Establish active execution"}
// Enter Running and evaluate both children; owner Result stays NotEvaluated until finalization.
FSteps[3].ExpectedState := E_State.Running;
FSteps[3].ExpectedResult := E_Result.NotEvaluated;
FSteps[3].ExpectedReady := FALSE;
FSteps[3].ExpectedPassedCount := 2;
FSteps[3].ExpectedFailedCount := 0;
FSteps[3].ExpectedHookCount := 5;
FSteps[3].ExpectedHooks[1].Hook := E_LifecycleHook.Abort;
FSteps[3].ExpectedHooks[1].State := E_State.Running;
FSteps[3].ExpectedHooks[1].Enabled := FALSE;
FSteps[3].ExpectedHooks[2].Hook := E_LifecycleHook.Preparations;
FSteps[3].ExpectedHooks[2].State := E_State.Running;
FSteps[3].ExpectedHooks[2].Enabled := FALSE;
FSteps[3].ExpectedHooks[3].Hook := E_LifecycleHook.Tests;
FSteps[3].ExpectedHooks[3].State := E_State.Running;
FSteps[3].ExpectedHooks[3].Enabled := TRUE;
FSteps[3].ExpectedHooks[4].Hook := E_LifecycleHook.Assertions;
FSteps[3].ExpectedHooks[4].State := E_State.Running;
FSteps[3].ExpectedHooks[4].Enabled := TRUE;
FSteps[3].ExpectedHooks[5].Hook := E_LifecycleHook.Aggregate;
FSteps[3].ExpectedHooks[5].State := E_State.Running;
FSteps[3].ExpectedHooks[5].Enabled := TRUE;
{endregion}

{region "04 - Request Abort and hold cleanup"}
// Enter Aborting and keep cleanup open so a later cleanup error can be injected.
FSteps[4].RequestAbort := TRUE;
FSteps[4].AbortCompleted := FALSE;
FSteps[4].ExpectedState := E_State.Aborting;
FSteps[4].ExpectedResult := E_Result.Abort;
FSteps[4].ExpectedReady := FALSE;
FSteps[4].ExpectedPassedCount := 2;
FSteps[4].ExpectedFailedCount := 0;
FSteps[4].ExpectedHookCount := 5;
FSteps[4].ExpectedHooks[1].Hook := E_LifecycleHook.Abort;
FSteps[4].ExpectedHooks[1].State := E_State.Aborting;
FSteps[4].ExpectedHooks[1].Enabled := TRUE;
FSteps[4].ExpectedHooks[2].Hook := E_LifecycleHook.Preparations;
FSteps[4].ExpectedHooks[2].State := E_State.Aborting;
FSteps[4].ExpectedHooks[2].Enabled := FALSE;
FSteps[4].ExpectedHooks[3].Hook := E_LifecycleHook.Tests;
FSteps[4].ExpectedHooks[3].State := E_State.Aborting;
FSteps[4].ExpectedHooks[3].Enabled := FALSE;
FSteps[4].ExpectedHooks[4].Hook := E_LifecycleHook.Assertions;
FSteps[4].ExpectedHooks[4].State := E_State.Aborting;
FSteps[4].ExpectedHooks[4].Enabled := FALSE;
FSteps[4].ExpectedHooks[5].Hook := E_LifecycleHook.Aggregate;
FSteps[4].ExpectedHooks[5].State := E_State.Aborting;
FSteps[4].ExpectedHooks[5].Enabled := TRUE;
{endregion}

{region "05 - Escalate cleanup failure to Error"}
// Raise Error inside the active Abort hook; Error must dominate Abort.
// This hook enters Aborting, while subsequent hooks observe AbortingFromError.
FSteps[5].AbortError := TRUE;
FSteps[5].AbortCompleted := FALSE;
FSteps[5].ExpectedState := E_State.AbortingFromError;
FSteps[5].ExpectedResult := E_Result.Error;
FSteps[5].ExpectedReady := FALSE;
FSteps[5].ExpectedPassedCount := 2;
FSteps[5].ExpectedFailedCount := 0;
FSteps[5].ExpectedHookCount := 5;
FSteps[5].ExpectedHooks[1].Hook := E_LifecycleHook.Abort;
FSteps[5].ExpectedHooks[1].State := E_State.Aborting;
FSteps[5].ExpectedHooks[1].Enabled := TRUE;
FSteps[5].ExpectedHooks[2].Hook := E_LifecycleHook.Preparations;
FSteps[5].ExpectedHooks[2].State := E_State.AbortingFromError;
FSteps[5].ExpectedHooks[2].Enabled := FALSE;
FSteps[5].ExpectedHooks[3].Hook := E_LifecycleHook.Tests;
FSteps[5].ExpectedHooks[3].State := E_State.AbortingFromError;
FSteps[5].ExpectedHooks[3].Enabled := FALSE;
FSteps[5].ExpectedHooks[4].Hook := E_LifecycleHook.Assertions;
FSteps[5].ExpectedHooks[4].State := E_State.AbortingFromError;
FSteps[5].ExpectedHooks[4].Enabled := FALSE;
FSteps[5].ExpectedHooks[5].Hook := E_LifecycleHook.Aggregate;
FSteps[5].ExpectedHooks[5].State := E_State.AbortingFromError;
FSteps[5].ExpectedHooks[5].Enabled := TRUE;
{endregion}

{region "06 - Acknowledge error cleanup"}
// Acknowledge cleanup on the next call; finalization must retain Error, not downgrade to Abort.
FSteps[6].ExpectedState := E_State.Completing;
FSteps[6].ExpectedResult := E_Result.Error;
FSteps[6].ExpectedReady := FALSE;
FSteps[6].ExpectedPassedCount := 2;
FSteps[6].ExpectedFailedCount := 0;
FSteps[6].ExpectedHookCount := 5;
FSteps[6].ExpectedHooks[1].Hook := E_LifecycleHook.Abort;
FSteps[6].ExpectedHooks[1].State := E_State.AbortingFromError;
FSteps[6].ExpectedHooks[1].Enabled := TRUE;
FSteps[6].ExpectedHooks[2].Hook := E_LifecycleHook.Preparations;
FSteps[6].ExpectedHooks[2].State := E_State.Completing;
FSteps[6].ExpectedHooks[2].Enabled := FALSE;
FSteps[6].ExpectedHooks[3].Hook := E_LifecycleHook.Tests;
FSteps[6].ExpectedHooks[3].State := E_State.Completing;
FSteps[6].ExpectedHooks[3].Enabled := FALSE;
FSteps[6].ExpectedHooks[4].Hook := E_LifecycleHook.Assertions;
FSteps[6].ExpectedHooks[4].State := E_State.Completing;
FSteps[6].ExpectedHooks[4].Enabled := FALSE;
FSteps[6].ExpectedHooks[5].Hook := E_LifecycleHook.Aggregate;
FSteps[6].ExpectedHooks[5].State := E_State.Completing;
FSteps[6].ExpectedHooks[5].Enabled := TRUE;
{endregion}

{region "07 - Observe terminal Error"}
// The following call reaches Completed; only aggregation remains in the recorded processing
// hooks.
FSteps[7].ExpectedState := E_State.Completed;
FSteps[7].ExpectedResult := E_Result.Error;
FSteps[7].ExpectedReady := FALSE;
FSteps[7].ExpectedPassedCount := 2;
FSteps[7].ExpectedFailedCount := 0;
FSteps[7].ExpectedHookCount := 1;
FSteps[7].ExpectedHooks[1].Hook := E_LifecycleHook.Aggregate;
FSteps[7].ExpectedHooks[1].State := E_State.Completed;
FSteps[7].ExpectedHooks[1].Enabled := TRUE;
{endregion}
END_METHOD

END_FUNCTION_BLOCK

// ---- SelfTests/TestCases/TestSuite_TestCaseLifecycle/Test_LifecycleAbortTimeout.TcPOU
{region 'Documentation'}
(*!
<summary>Withholds CompleteAbort and verifies timeout finalization with the latched Abort timeout flag.</summary>
*)
{endregion}
FUNCTION_BLOCK Test_LifecycleAbortTimeout EXTENDS TestCaseLifecycleTestBase

SUPER^();

{region 'Documentation'}
(*!
<summary>Defines explicit exceptional-path stimuli and contract-derived observations.</summary>
*)
{endregion}
METHOD PROTECTED ConfigureScenario
// Exercise the real cyclic timer; these checkpoints check the timeout path and retained flag,
// not an exact elapsed-time boundary. The outer Test Case timeout bounds a missing transition.
FSubjectPreparationCount := 0;
FSubjectTestCount := 1;
FStepCount := 12;
FSubjectConfig.AbortTimeout := T#50ms;

{region "01 - Reset to Idle"}
// Establish Idle through the parent Reset request; both child results must be cleared.
FSteps[1].RequestReset := TRUE;
FSteps[1].ExpectedState := E_State.Idle;
FSteps[1].ExpectedResult := E_Result.NotEvaluated;
FSteps[1].ExpectedReady := TRUE;
FSteps[1].ExpectedPassedCount := 0;
FSteps[1].ExpectedFailedCount := 0;
FSteps[1].ExpectedHookCount := 6;
FSteps[1].ExpectedHooks[1].Hook := E_LifecycleHook.Reset;
FSteps[1].ExpectedHooks[1].State := E_State.Reset;
FSteps[1].ExpectedHooks[1].Enabled := TRUE;
FSteps[1].ExpectedHooks[2].Hook := E_LifecycleHook.Abort;
FSteps[1].ExpectedHooks[2].State := E_State.Idle;
FSteps[1].ExpectedHooks[2].Enabled := FALSE;
FSteps[1].ExpectedHooks[3].Hook := E_LifecycleHook.Preparations;
FSteps[1].ExpectedHooks[3].State := E_State.Idle;
FSteps[1].ExpectedHooks[3].Enabled := FALSE;
FSteps[1].ExpectedHooks[4].Hook := E_LifecycleHook.Tests;
FSteps[1].ExpectedHooks[4].State := E_State.Idle;
FSteps[1].ExpectedHooks[4].Enabled := FALSE;
FSteps[1].ExpectedHooks[5].Hook := E_LifecycleHook.Assertions;
FSteps[1].ExpectedHooks[5].State := E_State.Idle;
FSteps[1].ExpectedHooks[5].Enabled := FALSE;
FSteps[1].ExpectedHooks[6].Hook := E_LifecycleHook.Aggregate;
FSteps[1].ExpectedHooks[6].State := E_State.Idle;
FSteps[1].ExpectedHooks[6].Enabled := TRUE;
{endregion}

